--- program second_half_topPaint (robot ABB IRB 5500-27) ---
  Smooth(1)
  Set speed (1000.0 mm/s)
  Set Ref.: FrameTopPaint
  Set Tool: Paint gun
  Show Paint gun
  MoveJ 1 to (-680.86, -907.35, 967.38) mm, rotated rx -105.87 ry 21.86 rz 12.34 deg; joints [-6.464, -4.331, 30.186, -24.09, 51.501, -71.972, -33.04]
  MoveL 2 to (-680.86, -907.35, 967.38) mm, rotated rx -105.87 ry 21.86 rz 12.34 deg; joints [-6.464, -4.331, 30.186, -24.09, 51.501, -71.972, -33.04]
  MoveL 3 to (-711.37, -815.56, 942.01) mm, rotated rx -105.87 ry 21.86 rz 12.34 deg; joints [-10.668, -3.752, 30.735, -25.583, 48.262, -68.348, -33.04]
  MoveL 4 to (-711.37, -815.56, 942.01) mm, rotated rx -105.87 ry 21.86 rz 12.34 deg; joints [-10.668, -3.752, 30.735, -25.583, 48.262, -68.348, -33.04]
  Set speed (50.0 mm/s)
  MoveL 5 to (-723.88, -815.55, 955.73) mm, rotated rx -113.43 ry 35.95 rz 5.6 deg; joints [-9.665, -1.677, 29.706, -47.736, 72.372, -53.861, -33.04]
  MoveL 6 to (-737.5, -815.56, 968.17) mm, rotated rx -117.99 ry 31.14 rz 6.09 deg; joints [-11, -4.053, 28.612, -30.497, 55.555, -56.043, -33.04]
  MoveL 7 to (-752.19, -815.56, 979.36) mm, rotated rx -123.35 ry 26.63 rz 6.68 deg; joints [-13.045, -6.077, 27.151, -7.256, 36.064, -62.575, -33.04]
  MoveL 8 to (-767.89, -815.56, 989.32) mm, rotated rx -137.44 ry 37.1 rz -8.5 deg; joints [-11.723, -3.945, 24.767, -26.574, 60.815, -46.836, -33.04]
  MoveL 9 to (-784.28, -815.56, 997.94) mm, rotated rx -143.37 ry 31.77 rz -8.88 deg; joints [-14.072, -5.42, 22.852, -4.109, 43.017, -52.262, -33.04]
  MoveL 10 to (-800.88, -815.56, 1005.13) mm, rotated rx -160.16 ry 35.48 rz -30.34 deg; joints [-12.936, -2.465, 18.781, -17.366, 67.621, -42.158, -33.04]
  MoveL 11 to (-817.93, -815.56, 1011.14) mm, rotated rx -163.51 ry 29.4 rz -30.19 deg; joints [-15.139, -2.909, 16.546, 0.625, 55.012, -47.084, -33.04]
  MoveL 12 to (-835.41, -815.56, 1016.08) mm, rotated rx -166.27 ry 23.89 rz -30.04 deg; joints [-17.301, -2.699, 14.273, 18.529, 44.337, -54.274, -33.04]
  MoveL 13 to (-853.23, -815.56, 1019.98) mm, rotated rx -168.26 ry 19.06 rz -29.89 deg; joints [-19.167, -1.967, 12.063, 35.166, 36.001, -62.757, -33.04]
  MoveL 14 to (-876.49, -815.56, 1023.58) mm, rotated rx -175.04 ry 16.66 rz -50.25 deg; joints [-17.559, 3.114, 5.489, 8.811, 70.793, -51.29, -33.04]
  MoveL 15 to (-899.83, -815.56, 1025.72) mm, rotated rx -173.61 ry 13.04 rz -49.71 deg; joints [-18.535, 4.811, 2.72, 14.774, 69.055, -56.135, -33.04]
  MoveL 16 to (-923.23, -815.56, 1026.54) mm, rotated rx -171.44 ry 10.87 rz -49.25 deg; joints [-18.954, 6.702, 0.191, 17.247, 69.288, -60.212, -33.04]
  MoveL 17 to (-946.69, -815.56, 1026.19) mm, rotated rx -168.63 ry 9.9 rz -48.73 deg; joints [-18.93, 8.673, -2.078, 17.142, 70.618, -63.617, -33.04]
  MoveL 18 to (-970.21, -815.56, 1024.77) mm, rotated rx -165.25 ry 9.92 rz -48.01 deg; joints [-18.58, 10.662, -4.07, 15.251, 72.434, -66.538, -33.04]
  MoveL 19 to (-993.66, -815.56, 1022.37) mm, rotated rx -161.4 ry 10.72 rz -47 deg; joints [-18.006, 12.618, -5.747, 12.177, 74.323, -69.099, -33.04]
  MoveL 20 to (-1016.91, -815.56, 1019.13) mm, rotated rx -154.6 ry 3.88 rz -27.21 deg; joints [-20.046, 11.059, -3.932, 50.238, 41.644, -92.598, -33.04]
  MoveL 21 to (-1052.97, -815.56, 1012.53) mm, rotated rx -147.18 ry 4.39 rz -25.42 deg; joints [-18.692, 13.832, -5.844, 42.524, 45.231, -94.781, -33.04]
  MoveL 22 to (-1088.6, -815.56, 1004.28) mm, rotated rx -139.61 ry 5.07 rz -23.14 deg; joints [-17.477, 16.361, -7.122, 35.707, 47.402, -97.128, -33.04]
  MoveL 23 to (-1123.86, -815.56, 994.58) mm, rotated rx -132.39 ry 5.54 rz -20.58 deg; joints [-16.529, 18.641, -7.948, 30.174, 48.333, -99.549, -33.04]
  MoveL 24 to (-1158.78, -815.56, 983.54) mm, rotated rx -125.85 ry 5.63 rz -17.99 deg; joints [-15.878, 20.702, -8.533, 26.043, 48.294, -101.998, -33.04]
  MoveL 25 to (-1193.38, -815.56, 971.26) mm, rotated rx -120.15 ry 5.32 rz -15.55 deg; joints [-15.49, 22.587, -9.043, 23.251, 47.542, -104.469, -33.04]
  MoveL 26 to (-1227.05, -815.55, 958.05) mm, rotated rx -117.54 ry 22.59 rz -22.51 deg; joints [-13.683, 27.315, -10.358, -19.064, 74.787, -84.054, -33.04]
  MoveL 27 to (-1260.34, -815.56, 943.78) mm, rotated rx -113.27 ry 22.78 rz -19.28 deg; joints [-13.733, 28.84, -10.662, -21.178, 73.313, -84.803, -33.04]
  MoveL 28 to (-1293.64, -815.56, 929.57) mm, rotated rx -110.3 ry 24.42 rz -16.76 deg; joints [-13.802, 30.363, -10.975, -25.489, 73.688, -83.558, -33.04]
  MoveL 29 to (-1326.93, -815.55, 915.36) mm, rotated rx -110.75 ry 26.95 rz -16.83 deg; joints [-13.938, 32.012, -12.325, -29.467, 76.004, -81.006, -33.04]
  Set speed (1000.0 mm/s)
  MoveL 30 to (-1326.93, -815.55, 915.36) mm, rotated rx -110.75 ry 26.95 rz -16.83 deg; joints [-13.938, 32.012, -12.325, -29.467, 76.004, -81.006, -33.04]
  MoveL 31 to (-1338.64, -909.72, 946.94) mm, rotated rx -108.61 ry 8.09 rz -9.79 deg; joints [-12.86, 29.886, -14.209, 10.126, 49.766, -104.847, -33.04]
  Set speed (1000.0 mm/s)
  MoveL 32 to (-1427.54, -801.91, 1165.8) mm, rotated rx -168.37 ry 26.91 rz -49.4 deg; joints [-18.397, 27.533, -26.297, -2.238, 74.394, -59.791, -33.04]
  MoveL 33 to (-1441.08, -755.13, 1078.46) mm, rotated rx -168.37 ry 26.91 rz -49.4 deg; joints [-19.651, 28.149, -23.955, -2.229, 72.544, -56.455, -33.04]
  MoveL 34 to (-1441.08, -755.13, 1078.46) mm, rotated rx -168.37 ry 26.91 rz -49.4 deg; joints [-19.651, 28.149, -23.955, -2.229, 72.544, -56.455, -33.04]
  Set speed (50.0 mm/s)
  MoveL 35 to (-1392.85, -755.13, 1070.73) mm, rotated rx -167.45 ry 26.52 rz -49.02 deg; joints [-19.416, 26.202, -21.042, -2.719, 73.023, -56.398, -33.04]
  MoveL 36 to (-1344.51, -755.13, 1064.62) mm, rotated rx -166.39 ry 26.02 rz -48.59 deg; joints [-19.179, 24.323, -18.348, -2.991, 73.454, -56.694, -33.04]
  MoveL 37 to (-1296.05, -755.13, 1060.31) mm, rotated rx -165.14 ry 25.36 rz -48.07 deg; joints [-18.944, 22.516, -15.888, -2.97, 73.811, -57.435, -33.04]
  MoveL 38 to (-1247.5, -755.13, 1057.45) mm, rotated rx -163.92 ry 24.63 rz -47.58 deg; joints [-18.714, 20.718, -13.548, -2.801, 74.124, -58.304, -33.04]
  MoveL 39 to (-1198.88, -755.13, 1055.53) mm, rotated rx -162.66 ry 23.79 rz -47.07 deg; joints [-18.49, 18.954, -11.35, -2.42, 74.383, -59.409, -33.04]
  MoveL 40 to (-1154.65, -755.13, 1054.25) mm, rotated rx -161.47 ry 22.9 rz -46.6 deg; joints [-18.296, 17.383, -9.469, -1.877, 74.573, -60.622, -33.04]
  MoveL 41 to (-1110.41, -755.13, 1053.12) mm, rotated rx -160.23 ry 21.86 rz -46.13 deg; joints [-18.116, 15.849, -7.702, -1.119, 74.72, -62.054, -33.04]
  MoveL 42 to (-1066.18, -755.13, 1051.84) mm, rotated rx -158.93 ry 20.61 rz -45.66 deg; joints [-17.96, 14.367, -6.063, -0.094, 74.823, -63.754, -33.04]
  MoveL 43 to (-1021.98, -755.13, 1050.14) mm, rotated rx -155.56 ry 16.38 rz -27.11 deg; joints [-20.211, 7.807, 1.212, 35.102, 38.519, -76.601, -33.04]
  MoveL 44 to (-977.83, -755.13, 1047.71) mm, rotated rx -167.34 ry 20.31 rz -48.51 deg; joints [-18.414, 8.637, -0.031, 2.711, 72.736, -56.241, -33.04]
  MoveL 45 to (-933.79, -755.13, 1044.23) mm, rotated rx -172.03 ry 17.59 rz -49.64 deg; joints [-19.417, 5.728, 2.312, 9.306, 68.998, -54.431, -33.04]
  MoveL 46 to (-889.96, -755.13, 1039.39) mm, rotated rx -176.35 ry 15.79 rz -50.43 deg; joints [-20.284, 2.79, 5.029, 14.554, 65.44, -52.144, -33.04]
  MoveL 47 to (-859.98, -755.13, 1035.09) mm, rotated rx -179.05 ry 15.23 rz -50.85 deg; joints [-20.714, 0.773, 7.104, 16.981, 63.333, -50.184, -33.04]
  MoveL 48 to (-830.15, -755.13, 1029.86) mm, rotated rx 178.5 ry 15.31 rz -51.25 deg; joints [-20.935, -1.226, 9.339, 18.054, 61.765, -47.765, -33.04]
  MoveL 49 to (-800.49, -755.13, 1023.59) mm, rotated rx 176.32 ry 16.12 rz -51.7 deg; joints [-20.879, -3.182, 11.724, 17.357, 61.061, -44.748, -33.04]
  MoveL 50 to (-771.02, -755.13, 1016.11) mm, rotated rx 174.42 ry 17.73 rz -52.29 deg; joints [-20.476, -5.053, 14.244, 14.483, 61.629, -41.047, -33.04]
  MoveL 51 to (-746.27, -755.13, 1008.74) mm, rotated rx 173.04 ry 19.75 rz -52.97 deg; joints [-19.815, -6.52, 16.467, 10.081, 63.46, -37.399, -33.04]
  MoveL 52 to (-721.93, -755.13, 1000.39) mm, rotated rx 171.85 ry 22.37 rz -53.89 deg; joints [-18.839, -7.804, 18.74, 3.824, 66.801, -33.461, -33.04]
  MoveL 53 to (-698.07, -755.13, 991) mm, rotated rx 170.81 ry 25.58 rz -55.13 deg; joints [-17.554, -8.832, 21.041, -4.204, 71.863, -29.519, -33.04]
  MoveL 54 to (-674.71, -755.13, 980.5) mm, rotated rx -178.47 ry 30.85 rz -33.67 deg; joints [-19.518, -13.327, 26.774, 8.833, 42.793, -34.507, -33.04]
  MoveL 55 to (-651.88, -755.13, 968.81) mm, rotated rx -177.42 ry 35.05 rz -34.68 deg; joints [-17.437, -13.741, 29.013, -6.651, 53.844, -28.419, -33.04]
  MoveL 56 to (-629.61, -755.13, 955.87) mm, rotated rx -176.18 ry 39.58 rz -35.92 deg; joints [-15.275, -13.645, 31.207, -21.324, 65.847, -24.476, -33.04]
  MoveL 57 to (-609.19, -755.13, 942.47) mm, rotated rx -157.46 ry 39.23 rz -11.27 deg; joints [-17.521, -17.024, 35.308, -13.254, 41.312, -30.381, -33.04]
  MoveL 58 to (-589.56, -755.13, 927.98) mm, rotated rx -153.88 ry 43.02 rz -11.42 deg; joints [-15.133, -16.253, 37.231, -29.816, 56.214, -26.857, -33.04]
  MoveL 59 to (-570.79, -755.13, 912.43) mm, rotated rx -150.35 ry 46.8 rz -11.58 deg; joints [-13.086, -14.971, 38.921, -43.447, 70.123, -26.03, -33.04]
  MoveL 60 to (-552.87, -755.13, 895.83) mm, rotated rx -132.12 ry 37.38 rz 9.39 deg; joints [-15.418, -17.926, 41.46, -31.974, 44.911, -34.545, -33.04]
  MoveL 61 to (-535.98, -755.13, 878.3) mm, rotated rx -128.2 ry 40.11 rz 9.17 deg; joints [-13.411, -16.317, 42.937, -45.251, 59.152, -33.515, -33.04]
  MoveL 62 to (-519.26, -755.12, 858.88) mm, rotated rx -124.45 ry 42.99 rz 8.96 deg; joints [-11.739, -14.257, 44.196, -56.795, 72.787, -34.124, -33.04]
  MoveL 63 to (-503.73, -755.13, 838.65) mm, rotated rx -114.08 ry 28.02 rz 20.35 deg; joints [-13.853, -17.337, 45.471, -36.435, 43.409, -46.335, -33.04]
  MoveL 64 to (-489.34, -755.13, 817.63) mm, rotated rx -111.22 ry 30.33 rz 19.47 deg; joints [-12.23, -15.335, 46.617, -48.302, 56.678, -44.847, -33.04]
  MoveL 65 to (-476.03, -755.13, 795.85) mm, rotated rx -108.72 ry 32.65 rz 18.71 deg; joints [-10.971, -13.136, 47.527, -57.964, 68.476, -44.674, -33.04]
  MoveL 66 to (-463.75, -755.13, 773.36) mm, rotated rx -104.02 ry 15.61 rz 23.88 deg; joints [-13.073, -16.444, 47.716, -24.573, 33.094, -63.727, -33.04]
  MoveL 67 to (-452.46, -755.13, 750.19) mm, rotated rx -102.19 ry 17.65 rz 22.76 deg; joints [-11.641, -14.473, 48.652, -37.695, 45.898, -59.342, -33.04]
  Set speed (1000.0 mm/s)
  MoveL 68 to (-452.46, -755.13, 750.19) mm, rotated rx -102.19 ry 17.65 rz 22.76 deg; joints [-11.641, -14.473, 48.652, -37.695, 45.898, -59.342, -33.04]
  MoveL 69 to (-408.75, -842.79, 770.31) mm, rotated rx -102.19 ry 17.65 rz 22.76 deg; joints [-5.982, -16.094, 48.843, -32.575, 47.942, -65.004, -33.04]
  Set speed (1000.0 mm/s)
  MoveL 70 to (-280.85, -767.56, 751.15) mm, rotated rx -114.97 ry 33.92 rz 24.38 deg; joints [-10.377, -28.704, 57.94, -50.266, 54.482, -37.789, -33.04]
  MoveL 71 to (-339.72, -694.7, 716.13) mm, rotated rx -114.97 ry 33.92 rz 24.38 deg; joints [-16.491, -24.096, 57.105, -61.18, 58.103, -29.538, -33.04]
  MoveL 72 to (-339.72, -694.7, 716.13) mm, rotated rx -114.97 ry 33.92 rz 24.38 deg; joints [-16.491, -24.096, 57.105, -61.18, 58.103, -29.538, -33.04]
  Set speed (50.0 mm/s)
  MoveL 73 to (-357.11, -694.7, 743.86) mm, rotated rx -117.94 ry 32.09 rz 25.15 deg; joints [-18.606, -26.389, 55.654, -51.693, 45.003, -28.551, -33.04]
  MoveL 74 to (-375.74, -694.69, 770.58) mm, rotated rx -130.67 ry 46.61 rz 11.02 deg; joints [-15.598, -23.039, 54.114, -63.974, 72.081, -20.66, -33.04]
  MoveL 75 to (-395.64, -694.7, 796.31) mm, rotated rx -134.35 ry 44.15 rz 11.08 deg; joints [-17.761, -25.145, 52.527, -53.816, 58.424, -18.794, -33.04]
  MoveL 76 to (-416.85, -694.7, 820.98) mm, rotated rx -138.3 ry 41.66 rz 11.13 deg; joints [-20.283, -26.646, 50.605, -42.162, 44.019, -18.14, -33.04]
  MoveL 77 to (-439.4, -694.7, 844.57) mm, rotated rx -159.64 ry 49.05 rz -13.25 deg; joints [-17.084, -23.648, 47.731, -45.094, 65.338, -13.723, -33.04]
  MoveL 78 to (-462.87, -694.7, 866.64) mm, rotated rx -162.58 ry 45.48 rz -12.83 deg; joints [-19.593, -24.599, 45.602, -31.764, 50.861, -14.485, -33.04]
  MoveL 79 to (-487.43, -694.7, 887.42) mm, rotated rx 175.77 ry 43.79 rz -39.75 deg; joints [-16.92, -21.228, 41.257, -31.131, 70.359, -12.811, -33.04]
  MoveL 80 to (-513.03, -694.7, 906.91) mm, rotated rx 175.37 ry 39.79 rz -37.93 deg; joints [-19.194, -21.396, 38.943, -17.947, 57.935, -15.44, -33.04]
  MoveL 81 to (-539.61, -694.7, 925.1) mm, rotated rx 174.96 ry 35.98 rz -36.42 deg; joints [-21.423, -21.016, 36.518, -3.67, 46.106, -20.168, -33.04]
  MoveL 82 to (-567.52, -694.7, 942.26) mm, rotated rx 162.99 ry 28.48 rz -57.97 deg; joints [-19.195, -16.589, 30.728, -8.728, 70.789, -18.654, -33.04]
  MoveL 83 to (-596.05, -694.71, 958.02) mm, rotated rx 164.29 ry 25.51 rz -56.36 deg; joints [-20.66, -15.521, 28.236, -0.029, 64.448, -22.61, -33.04]
  MoveL 84 to (-625.13, -694.71, 972.48) mm, rotated rx 165.62 ry 23.02 rz -55.12 deg; joints [-21.799, -14.167, 25.764, 7.202, 59.845, -26.748, -33.04]
  MoveL 85 to (-654.73, -694.71, 985.73) mm, rotated rx 167.01 ry 21.02 rz -54.2 deg; joints [-22.603, -12.611, 23.335, 12.74, 56.867, -30.707, -33.04]
  MoveL 86 to (-684.8, -694.71, 997.88) mm, rotated rx 168.52 ry 19.53 rz -53.53 deg; joints [-23.088, -10.915, 20.962, 16.48, 55.343, -34.23, -33.04]
  MoveL 87 to (-715.3, -694.71, 1009.03) mm, rotated rx 170.16 ry 18.56 rz -53.05 deg; joints [-23.288, -9.129, 18.656, 18.478, 55.039, -37.199, -33.04]
  MoveL 88 to (-746.19, -694.71, 1019.28) mm, rotated rx 171.94 ry 18.1 rz -52.71 deg; joints [-23.247, -7.286, 16.425, 18.902, 55.71, -39.601, -33.04]
  MoveL 89 to (-790.01, -694.71, 1032.3) mm, rotated rx 171.82 ry 18.31 rz -52.78 deg; joints [-23.382, -5.469, 14.353, 18.926, 55.572, -39.688, -33.04]
  MoveL 90 to (-834.27, -694.71, 1044) mm, rotated rx -164.38 ry 12.66 rz -47.66 deg; joints [-21.172, 3.673, 3.763, 15.498, 67.78, -65.474, -33.04]
  MoveL 91 to (-878.76, -694.71, 1054.62) mm, rotated rx -165.86 ry 14.3 rz -47.99 deg; joints [-21.21, 4.9, 2.353, 14.26, 67.353, -63.309, -33.04]
  MoveL 92 to (-923.43, -694.71, 1064.45) mm, rotated rx -167.05 ry 15.38 rz -48.3 deg; joints [-21.336, 6.309, 0.654, 13.66, 66.935, -61.91, -33.04]
  MoveL 93 to (-968.22, -694.71, 1073.75) mm, rotated rx -168.04 ry 16.15 rz -48.56 deg; joints [-21.499, 7.83, -1.235, 13.422, 66.525, -60.996, -33.04]
  MoveL 94 to (-1026.95, -694.71, 1085.57) mm, rotated rx -169.1 ry 16.87 rz -48.86 deg; joints [-21.736, 9.93, -3.917, 13.442, 66.008, -60.295, -33.04]
  MoveL 95 to (-1085.65, -694.71, 1097.49) mm, rotated rx -170.03 ry 17.43 rz -49.12 deg; joints [-21.979, 12.104, -6.785, 13.695, 65.517, -59.971, -33.04]
  MoveL 96 to (-1144.22, -694.71, 1110.04) mm, rotated rx -170.86 ry 17.87 rz -49.36 deg; joints [-22.222, 14.329, -9.82, 14.113, 65.054, -59.935, -33.04]
  MoveL 97 to (-1179.59, -694.71, 1109.54) mm, rotated rx -170.86 ry 17.87 rz -49.36 deg; joints [-22.351, 15.89, -11.706, 14.449, 64.884, -60.342, -33.04]
  MoveL 98 to (-1214.81, -694.71, 1107.82) mm, rotated rx -170.86 ry 17.87 rz -49.36 deg; joints [-22.474, 17.461, -13.593, 14.773, 64.725, -60.738, -33.04]
  MoveL 99 to (-1249.9, -694.71, 1104.91) mm, rotated rx -170.86 ry 17.87 rz -49.36 deg; joints [-22.592, 19.043, -15.485, 15.086, 64.575, -61.127, -33.04]
  MoveL 100 to (-1284.86, -694.71, 1100.85) mm, rotated rx -170.86 ry 17.87 rz -49.36 deg; joints [-22.705, 20.637, -17.385, 15.39, 64.435, -61.509, -33.04]
  MoveL 101 to (-1321.33, -694.71, 1095.39) mm, rotated rx -170.86 ry 17.87 rz -49.36 deg; joints [-22.819, 22.322, -19.388, 15.7, 64.298, -61.906, -33.04]
  MoveL 102 to (-1357.66, -694.71, 1088.73) mm, rotated rx -170.86 ry 17.87 rz -49.36 deg; joints [-22.928, 24.024, -21.407, 16.001, 64.172, -62.301, -33.04]
  MoveL 103 to (-1393.86, -694.71, 1080.88) mm, rotated rx -170.86 ry 17.87 rz -49.36 deg; joints [-23.032, 25.746, -23.447, 16.297, 64.055, -62.698, -33.04]
  Set speed (1000.0 mm/s)
  MoveL 104 to (-1393.86, -694.71, 1080.88) mm, rotated rx -170.86 ry 17.87 rz -49.36 deg; joints [-23.032, 25.746, -23.447, 16.297, 64.055, -62.698, -33.04]
  MoveL 105 to (-1386.19, -728.04, 1174.85) mm, rotated rx -170.86 ry 17.87 rz -49.36 deg; joints [-22.138, 25.351, -26.342, 16.111, 66.402, -66.107, -33.04]
  Set speed (1000.0 mm/s)
  MoveL 106 to (-1383.57, -648.28, 1177.84) mm, rotated rx -164.63 ry -10.56 rz -30.24 deg; joints [-29.593, 31.056, -38.749, 68.964, 56.594, -115.064, -33.04]
  MoveL 107 to (-1354.96, -634.29, 1083.04) mm, rotated rx -162.02 ry -4.77 rz -49.56 deg; joints [-27.513, 32.255, -36.738, 33.77, 75.893, -92.359, -33.04]
  MoveL 108 to (-1354.96, -634.29, 1083.04) mm, rotated rx -162.02 ry -4.77 rz -49.56 deg; joints [-27.513, 32.255, -36.738, 33.77, 75.893, -92.359, -33.04]
  Set speed (50.0 mm/s)
  MoveL 109 to (-1316.03, -634.28, 1090.58) mm, rotated rx -162.02 ry -4.77 rz -49.56 deg; joints [-27.496, 30.204, -34.071, 34.005, 75.314, -91.786, -33.04]
  MoveL 110 to (-1276.87, -634.28, 1096.8) mm, rotated rx -164.09 ry -4.88 rz -49.8 deg; joints [-27.831, 27.6, -30.819, 36.058, 73.417, -89.721, -33.04]
  MoveL 111 to (-1237.63, -634.28, 1101.65) mm, rotated rx -166.2 ry -4.97 rz -49.99 deg; joints [-28.188, 25.02, -27.61, 38.256, 71.356, -87.707, -33.04]
  MoveL 112 to (-1198.44, -634.28, 1105.09) mm, rotated rx -168.35 ry -5.02 rz -50.12 deg; joints [-28.564, 22.461, -24.431, 40.594, 69.113, -85.742, -33.04]
  MoveL 113 to (-1159.29, -634.28, 1107.12) mm, rotated rx -170.59 ry -4.99 rz -50.21 deg; joints [-28.959, 19.891, -21.234, 43.1, 66.607, -83.778, -33.04]
  MoveL 114 to (-1117.81, -634.28, 1107.7) mm, rotated rx -172.95 ry -4.89 rz -50.24 deg; joints [-29.388, 17.188, -17.865, 45.87, 63.758, -81.788, -33.04]
  MoveL 115 to (-1076.38, -634.28, 1106.64) mm, rotated rx -175.36 ry -4.66 rz -50.22 deg; joints [-29.827, 14.475, -14.468, 48.789, 60.627, -79.838, -33.04]
  MoveL 116 to (-1035, -634.28, 1103.91) mm, rotated rx -177.81 ry -4.29 rz -50.16 deg; joints [-30.273, 11.746, -11.032, 51.858, 57.195, -77.929, -33.04]
  MoveL 117 to (-993.67, -634.28, 1099.48) mm, rotated rx 179.68 ry -3.75 rz -50.05 deg; joints [-30.726, 8.988, -7.535, 55.102, 53.417, -76.051, -33.04]
  MoveL 118 to (-952.39, -634.28, 1093.3) mm, rotated rx 177.08 ry -3.02 rz -49.91 deg; joints [-31.187, 6.183, -3.95, 58.575, 49.223, -74.195, -33.04]
  MoveL 119 to (-911.16, -634.28, 1085.32) mm, rotated rx 170.97 ry -0.42 rz -49.61 deg; joints [-32.081, 1.909, 1.768, 66.623, 38.914, -70.262, -33.04]
  MoveL 120 to (-870.06, -634.28, 1072.26) mm, rotated rx 161.64 ry 24.15 rz -56.14 deg; joints [-25.915, -5.114, 14.971, 12.913, 51.726, -25.277, -33.04]
  MoveL 121 to (-829.03, -634.28, 1058.97) mm, rotated rx 161.64 ry 24.15 rz -56.14 deg; joints [-25.807, -6.839, 17.044, 12.396, 52.013, -24.786, -33.04]
  MoveL 122 to (-788.13, -634.28, 1045.27) mm, rotated rx 161.64 ry 24.15 rz -56.14 deg; joints [-25.693, -8.569, 19.094, 11.9, 52.305, -24.332, -33.04]
  MoveL 123 to (-747.44, -634.28, 1031) mm, rotated rx 161.64 ry 24.15 rz -56.14 deg; joints [-25.573, -10.301, 21.124, 11.421, 52.602, -23.909, -33.04]
  MoveL 124 to (-707.08, -634.28, 1015.99) mm, rotated rx 161.64 ry 24.15 rz -56.14 deg; joints [-25.446, -12.03, 23.135, 10.949, 52.909, -23.506, -33.04]
  MoveL 125 to (-667.17, -634.28, 1000.09) mm, rotated rx 161.64 ry 24.15 rz -56.14 deg; joints [-25.312, -13.749, 25.129, 10.477, 53.228, -23.113, -33.04]
  MoveL 126 to (-627.79, -634.28, 983.13) mm, rotated rx 161.64 ry 24.15 rz -56.14 deg; joints [-25.169, -15.454, 27.11, 9.996, 53.562, -22.721, -33.04]
  MoveL 127 to (-589.03, -634.28, 964.94) mm, rotated rx 161.64 ry 24.15 rz -56.14 deg; joints [-25.018, -17.14, 29.081, 9.495, 53.916, -22.317, -33.04]
  MoveL 128 to (-521.38, -634.28, 928.72) mm, rotated rx 160.54 ry 25.2 rz -56.78 deg; joints [-24.397, -20.285, 33.162, 5.492, 56.262, -19.182, -33.04]
  MoveL 129 to (-488.54, -634.28, 908.62) mm, rotated rx 159.09 ry 27.55 rz -58.21 deg; joints [-23.17, -21.751, 35.826, -2.329, 61.681, -14.851, -33.04]
  MoveL 130 to (-456.44, -634.28, 887.04) mm, rotated rx 157.59 ry 30.29 rz -60.07 deg; joints [-21.582, -22.904, 38.513, -11.425, 68.849, -10.813, -33.04]
  MoveL 131 to (-425.22, -634.28, 863.92) mm, rotated rx 170.2 ry 39.25 rz -38.62 deg; joints [-24.275, -27.281, 44.353, -11.924, 47.46, -10, -33.04]
  MoveL 132 to (-397.94, -634.28, 841.74) mm, rotated rx 170.15 ry 42.47 rz -40.29 deg; joints [-22.129, -27.683, 46.769, -24.269, 58.676, -6.356, -33.04]
  MoveL 133 to (-371.77, -634.27, 818.47) mm, rotated rx 170.03 ry 45.79 rz -42.27 deg; joints [-19.915, -27.569, 49.069, -35.693, 70.343, -4.4, -33.04]
  MoveL 134 to (-346.75, -634.28, 794.12) mm, rotated rx -166.97 ry 48.65 rz -13.97 deg; joints [-23.649, -30.931, 53.337, -40.952, 52.991, -3.509, -33.04]
  MoveL 135 to (-322.86, -634.28, 768.67) mm, rotated rx -164.78 ry 51.68 rz -14.53 deg; joints [-21.227, -30.129, 55.493, -51.709, 65.924, -3.715, -33.04]
  MoveL 136 to (-300.1, -634.28, 742.13) mm, rotated rx -141.36 ry 45.05 rz 12.36 deg; joints [-25.779, -33.162, 58.341, -56.228, 47.993, -3.726, -33.04]
  MoveL 137 to (-278.48, -634.28, 714.5) mm, rotated rx -137.94 ry 47.13 rz 12.43 deg; joints [-23.334, -31.875, 60.333, -64.364, 60.071, -6.057, -33.04]
  MoveL 138 to (-257.97, -634.28, 685.8) mm, rotated rx -123.43 ry 33.52 rz 29.26 deg; joints [-27.848, -34.937, 61.807, -64.029, 38.79, -8.276, -33.04]
  Set speed (1000.0 mm/s)
  MoveL 139 to (-257.97, -634.28, 685.8) mm, rotated rx -123.43 ry 33.52 rz 29.26 deg; joints [-27.848, -34.937, 61.807, -64.029, 38.79, -8.276, -33.04]
  MoveL 140 to (-190.63, -692.21, 731.73) mm, rotated rx -134.65 ry 49.19 rz 12.51 deg; joints [-15.298, -37.261, 63.293, -59.641, 65.012, -17.041, -33.04]
  Set speed (1000.0 mm/s)
  MoveL 141 to (-122.9, -618.87, 712.66) mm, rotated rx -142.88 ry 47.91 rz 13.38 deg; joints [-29.119, -48.176, 66.475, -50.842, 38.175, -0.586, -33.04]
  MoveL 142 to (-194.43, -573.85, 659.22) mm, rotated rx -142.88 ry 47.91 rz 13.38 deg; joints [-32.599, -38.02, 65.244, -72.969, 55.346, 9.693, -33.04]
  MoveL 143 to (-194.43, -573.85, 659.22) mm, rotated rx -142.88 ry 47.91 rz 13.38 deg; joints [-32.599, -38.02, 65.244, -72.969, 55.346, 9.693, -33.04]
  Set speed (50.0 mm/s)
  MoveL 144 to (-219.42, -573.85, 691.19) mm, rotated rx -168.5 ry 53.82 rz -15.6 deg; joints [-26.592, -35.485, 62.253, -59.133, 66.795, 5.859, -33.04]
  MoveL 145 to (-245.66, -573.85, 721.92) mm, rotated rx -170.35 ry 50.93 rz -14.9 deg; joints [-29.075, -36.259, 59.872, -49.532, 54.056, 6.877, -33.04]
  MoveL 146 to (-273.13, -573.85, 751.4) mm, rotated rx 165.69 ry 46.89 rz -44 deg; joints [-24.248, -33.143, 55.523, -38.026, 67.49, 3.047, -33.04]
  MoveL 147 to (-301.84, -573.85, 779.65) mm, rotated rx 166.16 ry 43.83 rz -41.85 deg; joints [-26.546, -33.105, 53.003, -26.934, 55.657, 1.11, -33.04]
  MoveL 148 to (-331.74, -573.84, 806.69) mm, rotated rx 152.1 ry 33.68 rz -63.59 deg; joints [-23.32, -29.086, 47.36, -20.418, 72.694, -1.696, -33.04]
  MoveL 149 to (-362.3, -573.85, 832.06) mm, rotated rx 153.68 ry 31.23 rz -61.45 deg; joints [-25.042, -28.271, 44.813, -11.519, 64.603, -4.897, -33.04]
  MoveL 150 to (-393.95, -573.85, 856.32) mm, rotated rx 155.14 ry 28.97 rz -59.69 deg; joints [-26.496, -27.094, 42.224, -3.137, 57.77, -8.726, -33.04]
  MoveL 151 to (-426.44, -573.85, 879.33) mm, rotated rx 155.14 ry 28.97 rz -59.69 deg; joints [-26.613, -25.628, 40.437, -2.635, 57.395, -9.123, -33.04]
  MoveL 152 to (-459.61, -573.85, 901.11) mm, rotated rx 155.14 ry 28.97 rz -59.69 deg; joints [-26.721, -24.133, 38.65, -2.172, 57.051, -9.487, -33.04]
  MoveL 153 to (-499.91, -573.85, 925.56) mm, rotated rx 155.14 ry 28.97 rz -59.69 deg; joints [-26.84, -22.326, 36.52, -1.659, 56.673, -9.893, -33.04]
  MoveL 154 to (-541.01, -573.85, 948.56) mm, rotated rx 155.14 ry 28.97 rz -59.69 deg; joints [-26.95, -20.496, 34.383, -1.173, 56.32, -10.28, -33.04]
  MoveL 155 to (-582.81, -573.85, 970.29) mm, rotated rx 155.14 ry 28.97 rz -59.69 deg; joints [-27.051, -18.65, 32.237, -0.7, 55.985, -10.662, -33.04]
  MoveL 156 to (-625.21, -573.85, 990.93) mm, rotated rx 155.14 ry 28.97 rz -59.69 deg; joints [-27.145, -16.796, 30.078, -0.227, 55.66, -11.054, -33.04]
  MoveL 157 to (-668.11, -573.85, 1010.65) mm, rotated rx 155.14 ry 28.97 rz -59.69 deg; joints [-27.234, -14.939, 27.903, 0.257, 55.338, -11.465, -33.04]
  MoveL 158 to (-711.41, -573.85, 1029.64) mm, rotated rx 155.14 ry 28.97 rz -59.69 deg; joints [-27.317, -13.084, 25.708, 0.764, 55.014, -11.906, -33.04]
  MoveL 159 to (-748.06, -573.85, 1043.66) mm, rotated rx 157.61 ry 6.44 rz -70.97 deg; joints [-30.214, -6.982, 13.644, 24.862, 64.48, -31.395, -33.04]
  MoveL 160 to (-785.01, -573.85, 1056.24) mm, rotated rx 159.54 ry 6.06 rz -70.87 deg; joints [-30.059, -4.756, 10.809, 24.468, 66.213, -33.972, -33.04]
  MoveL 161 to (-822.27, -573.85, 1067.4) mm, rotated rx 161.68 ry 5.81 rz -70.82 deg; joints [-29.825, -2.438, 7.89, 23.534, 68.351, -36.593, -33.04]
  MoveL 162 to (-859.82, -573.85, 1077.12) mm, rotated rx 163.93 ry 5.7 rz -70.8 deg; joints [-29.537, -0.058, 4.925, 22.194, 70.729, -39.212, -33.04]
  MoveL 163 to (-897.67, -573.85, 1085.42) mm, rotated rx 166.26 ry 5.73 rz -70.79 deg; joints [-29.212, 2.369, 1.93, 20.532, 73.248, -41.818, -33.04]
  MoveL 164 to (-935.15, -573.85, 1092.2) mm, rotated rx 171.31 ry 9.42 rz -50.91 deg; joints [-31.484, 1.113, 4.075, 53.364, 36.921, -59.511, -33.04]
  MoveL 165 to (-972.91, -573.85, 1097.61) mm, rotated rx 173.72 ry 8.88 rz -50.75 deg; joints [-31.012, 3.518, 1.087, 50.816, 40.223, -61.321, -33.04]
  MoveL 166 to (-1010.95, -573.85, 1101.66) mm, rotated rx 176.22 ry 8.44 rz -50.58 deg; joints [-30.529, 5.963, -1.923, 48.198, 43.461, -63.201, -33.04]
  MoveL 167 to (-1049.28, -573.85, 1104.34) mm, rotated rx 179.02 ry 8.02 rz -50.35 deg; joints [-30.017, 8.52, -5.057, 45.445, 46.81, -65.379, -33.04]
  MoveL 168 to (-1095.21, -573.85, 1105.76) mm, rotated rx 178.6 ry -0.8 rz -49.98 deg; joints [-32.096, 12.453, -11.192, 57.274, 48.606, -75.574, -33.04]
  MoveL 169 to (-1141.03, -573.85, 1105.26) mm, rotated rx -179.95 ry -2.76 rz -50.03 deg; joints [-32.127, 15.498, -15.21, 56.44, 52.134, -78.187, -33.04]
  MoveL 170 to (-1186.71, -573.85, 1102.88) mm, rotated rx -178.47 ry -4.6 rz -50.15 deg; joints [-32.125, 18.597, -19.315, 55.198, 55.858, -80.655, -33.04]
  MoveL 171 to (-1232.24, -573.85, 1098.69) mm, rotated rx -176.96 ry -6.34 rz -50.33 deg; joints [-32.096, 21.761, -23.526, 53.627, 59.732, -83.045, -33.04]
  MoveL 172 to (-1277.62, -573.85, 1092.71) mm, rotated rx -175.43 ry -7.97 rz -50.56 deg; joints [-32.044, 25.002, -27.87, 51.781, 63.733, -85.408, -33.04]
  MoveL 173 to (-1322.87, -573.85, 1084.99) mm, rotated rx -173.88 ry -9.5 rz -50.83 deg; joints [-31.971, 28.336, -32.379, 49.693, 67.845, -87.788, -33.04]
  Set speed (1000.0 mm/s)
  MoveL 174 to (-1322.87, -573.85, 1084.99) mm, rotated rx -173.88 ry -9.5 rz -50.83 deg; joints [-31.971, 28.336, -32.379, 49.693, 67.845, -87.788, -33.04]
  MoveL 175 to (-1341.5, -567.86, 1183.06) mm, rotated rx -173.88 ry -9.5 rz -50.83 deg; joints [-32.09, 29.766, -38.022, 47.112, 72.847, -91.048, -33.04]
  Set speed (1000.0 mm/s)
  MoveL 176 to (-1313.29, -509.41, 1185.2) mm, rotated rx -174 ry -7.96 rz -50.61 deg; joints [-33.45, 27.776, -35.021, 50.071, 68.116, -90.852, -33.04]
  MoveL 177 to (-1296.48, -513.43, 1086.71) mm, rotated rx -174 ry -7.96 rz -50.61 deg; joints [-33.386, 26.559, -29.695, 52.526, 63.238, -87.794, -33.04]
  MoveL 178 to (-1296.48, -513.43, 1086.71) mm, rotated rx -174 ry -7.96 rz -50.61 deg; joints [-33.386, 26.559, -29.695, 52.526, 63.238, -87.794, -33.04]
  Set speed (50.0 mm/s)
  MoveL 179 to (-1258.34, -513.43, 1092.62) mm, rotated rx -175.35 ry -6.81 rz -50.43 deg; joints [-33.519, 23.847, -26.066, 54.385, 59.91, -85.983, -33.04]
  MoveL 180 to (-1220.17, -513.43, 1097.33) mm, rotated rx -176.67 ry -5.59 rz -50.28 deg; joints [-33.643, 21.197, -22.544, 56.13, 56.627, -84.205, -33.04]
  MoveL 181 to (-1182, -513.43, 1100.83) mm, rotated rx -177.98 ry -4.32 rz -50.15 deg; joints [-33.757, 18.6, -19.111, 57.751, 53.389, -82.439, -33.04]
  MoveL 182 to (-1143.81, -513.43, 1103.09) mm, rotated rx -179.27 ry -2.98 rz -50.06 deg; joints [-33.861, 16.049, -15.756, 59.23, 50.207, -80.666, -33.04]
  MoveL 183 to (-1104.9, -513.43, 1104.12) mm, rotated rx 179.43 ry -1.55 rz -50 deg; joints [-33.953, 13.492, -12.406, 60.563, 47.035, -78.826, -33.04]
  MoveL 184 to (-1065.98, -513.43, 1103.84) mm, rotated rx 178.15 ry -0.05 rz -49.98 deg; joints [-34.03, 10.973, -9.113, 61.684, 43.954, -76.92, -33.04]
  MoveL 185 to (-1027.05, -513.43, 1102.23) mm, rotated rx 176.88 ry 1.52 rz -50.02 deg; joints [-34.089, 8.485, -5.869, 62.538, 40.995, -74.907, -33.04]
  MoveL 186 to (-988.09, -513.43, 1099.26) mm, rotated rx 175.63 ry 3.14 rz -50.1 deg; joints [-34.128, 6.029, -2.671, 63.054, 38.21, -72.742, -33.04]
  MoveL 187 to (-949.11, -513.43, 1094.89) mm, rotated rx 173.09 ry 2.63 rz -70.17 deg; joints [-31.467, 7.286, -4.699, 23.829, 75.046, -52.259, -33.04]
  MoveL 188 to (-910.16, -513.43, 1089.13) mm, rotated rx 171.34 ry 3.87 rz -70.35 deg; joints [-31.36, 4.857, -1.509, 23.346, 73.511, -49.275, -33.04]
  MoveL 189 to (-871.59, -513.43, 1081.99) mm, rotated rx 169.6 ry 5.16 rz -70.6 deg; joints [-31.216, 2.485, 1.618, 22.513, 72.252, -46.22, -33.04]
  MoveL 190 to (-833.49, -513.43, 1073.52) mm, rotated rx 170.67 ry 6.91 rz -70.89 deg; joints [-30.503, 1.119, 3.619, 18.651, 74.196, -45.432, -33.04]
  MoveL 191 to (-795.86, -513.42, 1063.72) mm, rotated rx 170.67 ry 6.91 rz -70.89 deg; joints [-30.541, -0.485, 5.598, 18.7, 73.934, -45.052, -33.04]
  MoveL 192 to (-758.7, -513.42, 1052.61) mm, rotated rx 170.67 ry 6.91 rz -70.89 deg; joints [-30.58, -2.064, 7.563, 18.747, 73.667, -44.66, -33.04]
  MoveL 193 to (-719.79, -513.42, 1039.41) mm, rotated rx 170.67 ry 6.91 rz -70.89 deg; joints [-30.622, -3.712, 9.635, 18.794, 73.376, -44.23, -33.04]
  MoveL 194 to (-681.4, -513.42, 1024.77) mm, rotated rx 149.35 ry 33.54 rz -64.1 deg; joints [-28.786, -14.613, 29.431, -12.165, 61.244, -1.134, -33.04]
  MoveL 195 to (-643.51, -513.42, 1008.71) mm, rotated rx 149.35 ry 33.54 rz -64.1 deg; joints [-28.764, -16.254, 31.317, -12.486, 61.457, -0.85, -33.04]
  MoveL 196 to (-606.12, -513.42, 991.24) mm, rotated rx 149.35 ry 33.54 rz -64.1 deg; joints [-28.739, -17.877, 33.204, -12.834, 61.689, -0.544, -33.04]
  MoveL 197 to (-569.22, -513.42, 972.38) mm, rotated rx 149.35 ry 33.54 rz -64.1 deg; joints [-28.71, -19.483, 35.094, -13.21, 61.943, -0.217, -33.04]
  MoveL 198 to (-532.8, -513.42, 952.19) mm, rotated rx 149.35 ry 33.54 rz -64.1 deg; joints [-28.678, -21.072, 36.988, -13.612, 62.219, 0.131, -33.04]
  MoveL 199 to (-494.06, -513.42, 930.04) mm, rotated rx 149.35 ry 33.54 rz -64.1 deg; joints [-28.642, -22.787, 39.005, -14.014, 62.5, 0.473, -33.04]
  MoveL 200 to (-455.86, -513.42, 907) mm, rotated rx 149.35 ry 33.54 rz -64.1 deg; joints [-28.602, -24.499, 41.014, -14.411, 62.782, 0.808, -33.04]
  MoveL 201 to (-418.28, -513.42, 882.95) mm, rotated rx 149.35 ry 33.54 rz -64.1 deg; joints [-28.559, -26.2, 43.015, -14.812, 63.073, 1.142, -33.04]
  MoveL 202 to (-381.55, -513.42, 857.89) mm, rotated rx 149.35 ry 33.54 rz -64.1 deg; joints [-28.512, -27.877, 45.002, -15.228, 63.379, 1.484, -33.04]
  MoveL 203 to (-345.76, -513.42, 831.75) mm, rotated rx 149.35 ry 33.54 rz -64.1 deg; joints [-28.459, -29.523, 46.975, -15.668, 63.708, 1.843, -33.04]
  MoveL 204 to (-314.11, -513.42, 807) mm, rotated rx 149.35 ry 33.54 rz -64.1 deg; joints [-28.405, -30.985, 48.757, -16.099, 64.034, 2.191, -33.04]
  MoveL 205 to (-283.33, -513.42, 781.26) mm, rotated rx 149.35 ry 33.54 rz -64.1 deg; joints [-28.344, -32.406, 50.529, -16.57, 64.394, 2.57, -33.04]
  MoveL 206 to (-253.47, -513.42, 754.49) mm, rotated rx 149.35 ry 33.54 rz -64.1 deg; joints [-28.276, -33.78, 52.291, -17.091, 64.796, 2.986, -33.04]
  MoveL 207 to (-224.56, -513.42, 726.64) mm, rotated rx 163.14 ry 44.09 rz -42.56 deg; joints [-32.78, -37.601, 57.608, -26.32, 48.349, 7.862, -33.04]
  MoveL 208 to (-196.62, -513.42, 697.69) mm, rotated rx 162.55 ry 46.6 rz -44.46 deg; joints [-30.825, -37.995, 60.084, -36.188, 58.754, 10.127, -33.04]
  MoveL 209 to (-169.68, -513.41, 667.6) mm, rotated rx 161.8 ry 49.16 rz -46.66 deg; joints [-28.72, -37.819, 62.447, -45.533, 69.707, 11.196, -33.04]
  MoveL 210 to (-143.76, -513.42, 636.4) mm, rotated rx -172.47 ry 53.81 rz -16.01 deg; joints [-35.203, -40.241, 66.55, -63.162, 60.486, 17.594, -33.04]
  Set speed (1000.0 mm/s)
  MoveL 211 to (-143.76, -513.42, 636.4) mm, rotated rx -172.47 ry 53.81 rz -16.01 deg; joints [-35.203, -40.241, 66.55, -63.162, 60.486, 17.594, -33.04]
  MoveL 212 to (-70.48, -548.09, 694.95) mm, rotated rx -172.47 ry 53.81 rz -16.01 deg; joints [-33.329, -51.45, 67.814, -42.441, 43.539, 7.598, -33.04]
  Set speed (1000.0 mm/s)
  MoveL 213 to (-47.33, -481.42, 695.34) mm, rotated rx 159.13 ry 33.45 rz -61.67 deg; joints [-28.24, -45.438, 58.516, -9.181, 62.09, -12.887, -33.04]
  MoveL 214 to (-103.12, -452.99, 617.38) mm, rotated rx 159.13 ry 33.45 rz -61.67 deg; joints [-30.271, -38.474, 58.619, -15.757, 63.787, -4.136, -33.04]
  MoveL 215 to (-103.12, -452.99, 617.38) mm, rotated rx 159.13 ry 33.45 rz -61.67 deg; joints [-30.271, -38.474, 58.619, -15.757, 63.787, -4.136, -33.04]
  Set speed (50.0 mm/s)
  MoveL 216 to (-129.63, -452.99, 647.84) mm, rotated rx 159.46 ry 32.42 rz -60.95 deg; joints [-31.139, -37.612, 56.614, -11.317, 59.8, -5.914, -33.04]
  MoveL 217 to (-157.02, -452.99, 677.33) mm, rotated rx 159.79 ry 31.39 rz -60.25 deg; joints [-31.935, -36.598, 54.586, -6.876, 56.029, -7.838, -33.04]
  MoveL 218 to (-185.27, -452.99, 705.85) mm, rotated rx 160.11 ry 30.37 rz -59.59 deg; joints [-32.662, -35.458, 52.538, -2.411, 52.449, -9.918, -33.04]
  MoveL 219 to (-214.36, -452.99, 733.45) mm, rotated rx 160.44 ry 29.34 rz -58.94 deg; joints [-33.323, -34.213, 50.473, 2.092, 49.041, -12.161, -33.04]
  MoveL 220 to (-244.27, -452.99, 760.14) mm, rotated rx 160.77 ry 28.31 rz -58.33 deg; joints [-33.921, -32.88, 48.394, 6.648, 45.791, -14.573, -33.04]
  MoveL 221 to (-274.41, -452.99, 785.51) mm, rotated rx 161.11 ry 27.29 rz -57.74 deg; joints [-34.461, -31.499, 46.334, 11.259, 42.685, -17.147, -33.04]
  MoveL 222 to (-305.25, -452.99, 810.1) mm, rotated rx 153.74 ry 18.56 rz -77.17 deg; joints [-30.62, -26.126, 40.435, -0.493, 73.404, -13.225, -33.04]
  MoveL 223 to (-336.79, -452.99, 833.9) mm, rotated rx 154.42 ry 17.71 rz -76.57 deg; joints [-31.073, -24.721, 38.309, 2.176, 71.615, -14.981, -33.04]
  MoveL 224 to (-368.96, -453, 857.01) mm, rotated rx 155.1 ry 16.86 rz -76 deg; joints [-31.48, -23.261, 36.157, 4.742, 70.014, -16.782, -33.04]
  MoveL 225 to (-404.17, -453, 882.18) mm, rotated rx 155.78 ry 16.03 rz -75.46 deg; joints [-31.839, -21.661, 33.813, 7.235, 68.609, -18.708, -33.04]
  MoveL 226 to (-439.94, -453, 906.27) mm, rotated rx 156.47 ry 15.2 rz -74.95 deg; joints [-32.155, -20.015, 31.452, 9.602, 67.397, -20.653, -33.04]
  MoveL 227 to (-476.31, -453, 929.21) mm, rotated rx 157.17 ry 14.38 rz -74.46 deg; joints [-32.431, -18.322, 29.073, 11.835, 66.371, -22.605, -33.04]
  MoveL 228 to (-513.31, -453, 950.92) mm, rotated rx 158.03 ry 13.49 rz -73.96 deg; joints [-32.688, -16.54, 26.603, 14.089, 65.495, -24.788, -33.04]
  MoveL 229 to (-550.97, -453, 971.36) mm, rotated rx 158.59 ry 12.77 rz -73.58 deg; joints [-32.872, -14.798, 24.252, 15.873, 64.864, -26.492, -33.04]
  MoveL 230 to (-589.32, -453, 990.48) mm, rotated rx 159.32 ry 11.98 rz -73.19 deg; joints [-33.041, -12.967, 21.806, 17.667, 64.371, -28.41, -33.04]
  MoveL 231 to (-628.38, -453, 1008.24) mm, rotated rx 160.05 ry 11.21 rz -72.82 deg; joints [-33.18, -11.091, 19.333, 19.305, 64.045, -30.306, -33.04]
  MoveL 232 to (-664.81, -453, 1023.29) mm, rotated rx 160.76 ry 10.39 rz -72.45 deg; joints [-33.338, -9.324, 17.001, 20.987, 63.721, -32.184, -33.04]
  MoveL 233 to (-701.87, -453, 1037.14) mm, rotated rx 162.46 ry 9.16 rz -71.92 deg; joints [-33.495, -7.196, 14.161, 22.931, 63.912, -35.396, -33.04]
  MoveL 234 to (-739.57, -453, 1049.77) mm, rotated rx 164.18 ry 7.94 rz -71.45 deg; joints [-33.615, -5.001, 11.257, 24.556, 64.428, -38.561, -33.04]
  MoveL 235 to (-777.69, -453, 1061.07) mm, rotated rx 165.9 ry 6.74 rz -71.06 deg; joints [-33.698, -2.752, 8.305, 25.839, 65.255, -41.646, -33.04]
  MoveL 236 to (-815.99, -453, 1070.98) mm, rotated rx 167.62 ry 5.56 rz -70.73 deg; joints [-33.747, -0.466, 5.322, 26.781, 66.362, -44.63, -33.04]
  MoveL 237 to (-854.43, -453, 1079.52) mm, rotated rx 169.34 ry 4.43 rz -70.47 deg; joints [-33.766, 1.856, 2.305, 27.399, 67.722, -47.521, -33.04]
  MoveL 238 to (-900.78, -453, 1087.97) mm, rotated rx 171.4 ry 3.13 rz -70.24 deg; joints [-33.754, 4.69, -1.366, 27.739, 69.649, -50.878, -33.04]
  MoveL 239 to (-947.34, -453, 1094.5) mm, rotated rx 173.45 ry 1.9 rz -70.08 deg; joints [-33.707, 7.575, -5.096, 27.674, 71.852, -54.123, -33.04]
  MoveL 240 to (-994.13, -453, 1099.1) mm, rotated rx 175.51 ry 0.75 rz -70 deg; joints [-33.63, 10.515, -8.894, 27.242, 74.29, -57.284, -33.04]
  MoveL 241 to (-1041.13, -453, 1101.84) mm, rotated rx 177.6 ry 0.53 rz -49.99 deg; joints [-36.072, 9.806, -7.417, 67.04, 38.997, -78.938, -33.04]
  MoveL 242 to (-1088.35, -453, 1102.7) mm, rotated rx 179.2 ry -1.1 rz -49.99 deg; joints [-35.854, 12.798, -11.311, 64.962, 42.987, -80.75, -33.04]
  MoveL 243 to (-1134.94, -453, 1101.72) mm, rotated rx -179.2 ry -2.62 rz -50.05 deg; joints [-35.628, 15.797, -15.224, 62.78, 46.942, -82.533, -33.04]
  MoveL 244 to (-1181.72, -453, 1098.96) mm, rotated rx -177.57 ry -4.06 rz -50.15 deg; joints [-35.394, 18.863, -19.243, 60.486, 50.92, -84.351, -33.04]
  MoveL 245 to (-1228.42, -453, 1094.44) mm, rotated rx -175.93 ry -5.41 rz -50.28 deg; joints [-35.153, 21.989, -23.363, 58.106, 54.896, -86.219, -33.04]
  MoveL 246 to (-1274.93, -453, 1088.2) mm, rotated rx -174.27 ry -6.67 rz -50.44 deg; joints [-34.907, 25.18, -27.599, 55.655, 58.86, -88.151, -33.04]
  Set speed (1000.0 mm/s)
  MoveL 247 to (-1274.93, -453, 1088.2) mm, rotated rx -174.27 ry -6.67 rz -50.44 deg; joints [-34.907, 25.18, -27.599, 55.655, 58.86, -88.151, -33.04]
  MoveL 248 to (-1289.99, -450.45, 1187.03) mm, rotated rx -174.27 ry -6.67 rz -50.44 deg; joints [-34.929, 26.223, -32.676, 53.244, 63.693, -91.018, -33.04]
  Set speed (1000.0 mm/s)
  MoveL 249 to (-1255.42, -331.41, 1189.89) mm, rotated rx -175.11 ry -4.63 rz -50.22 deg; joints [-38.135, 24.154, -29.471, 60.413, 55.333, -92.348, -33.04]
  MoveL 250 to (-1243.73, -332.14, 1090.58) mm, rotated rx -175.11 ry -4.63 rz -50.22 deg; joints [-38.165, 23.385, -24.764, 62.958, 50.412, -89.891, -33.04]
  MoveL 251 to (-1243.73, -332.14, 1090.58) mm, rotated rx -175.11 ry -4.63 rz -50.22 deg; joints [-38.165, 23.385, -24.764, 62.958, 50.412, -89.891, -33.04]
  Set speed (50.0 mm/s)
  MoveL 252 to (-1201.21, -332.15, 1094.93) mm, rotated rx -176.65 ry -3.73 rz -50.14 deg; joints [-38.536, 20.631, -21.12, 65.782, 46.768, -88.717, -33.04]
  MoveL 253 to (-1158.6, -332.15, 1097.96) mm, rotated rx -178.19 ry -2.77 rz -50.07 deg; joints [-38.914, 17.921, -17.55, 68.73, 43.002, -87.689, -33.04]
  MoveL 254 to (-1116.04, -332.15, 1099.62) mm, rotated rx -179.13 ry -1.53 rz -70.03 deg; joints [-36.795, 18.924, -19.528, 29.457, 75.984, -66.765, -33.04]
  MoveL 255 to (-1073.65, -332.15, 1099.95) mm, rotated rx 179.1 ry -1.01 rz -69.99 deg; joints [-37.103, 16.233, -16.048, 31.062, 73.295, -64.446, -33.04]
  MoveL 256 to (-1031.4, -332.15, 1098.89) mm, rotated rx 177.31 ry -0.43 rz -69.96 deg; joints [-37.409, 13.588, -12.643, 32.546, 70.635, -62.144, -33.04]
  MoveL 257 to (-989.29, -332.15, 1096.44) mm, rotated rx 175.53 ry 0.22 rz -69.96 deg; joints [-37.715, 10.985, -9.302, 33.9, 68.013, -59.843, -33.04]
  MoveL 258 to (-943.54, -332.15, 1092.18) mm, rotated rx 173.58 ry 0.98 rz -69.98 deg; joints [-38.048, 8.188, -5.721, 35.213, 65.21, -57.321, -33.04]
  MoveL 259 to (-897.97, -332.15, 1086.25) mm, rotated rx 171.63 ry 1.82 rz -70.05 deg; joints [-38.378, 5.43, -2.197, 36.335, 62.485, -54.768, -33.04]
  MoveL 260 to (-852.58, -332.15, 1078.61) mm, rotated rx 169.68 ry 2.72 rz -70.16 deg; joints [-38.706, 2.708, 1.279, 37.244, 59.857, -52.162, -33.04]
  MoveL 261 to (-807.39, -332.15, 1069.24) mm, rotated rx 167.72 ry 3.68 rz -70.32 deg; joints [-39.031, 0.018, 4.712, 37.912, 57.35, -49.481, -33.04]
  MoveL 262 to (-762.39, -332.14, 1058.13) mm, rotated rx 165.76 ry 4.69 rz -70.53 deg; joints [-39.352, -2.639, 8.108, 38.309, 54.997, -46.708, -33.04]
  MoveL 263 to (-717.61, -332.14, 1045.24) mm, rotated rx 163.81 ry 5.74 rz -70.81 deg; joints [-39.667, -5.262, 11.466, 38.403, 52.828, -43.823, -33.04]
  MoveL 264 to (-673.51, -332.14, 1030.7) mm, rotated rx 161.86 ry 6.83 rz -71.15 deg; joints [-39.972, -7.829, 14.761, 38.163, 50.897, -40.831, -33.04]
  MoveL 265 to (-630.2, -332.14, 1014.58) mm, rotated rx 159.94 ry 7.92 rz -71.56 deg; joints [-40.265, -10.331, 17.985, 37.57, 49.235, -37.729, -33.04]
  MoveL 266 to (-587.66, -332.14, 996.91) mm, rotated rx 158.04 ry 9.02 rz -72.03 deg; joints [-40.544, -12.769, 21.141, 36.613, 47.864, -34.509, -33.04]
  MoveL 267 to (-545.88, -332.14, 977.73) mm, rotated rx 156.17 ry 10.11 rz -72.56 deg; joints [-40.81, -15.145, 24.235, 35.29, 46.801, -31.171, -33.04]
  MoveL 268 to (-504.84, -332.14, 957.06) mm, rotated rx 154.31 ry 11.18 rz -73.15 deg; joints [-41.062, -17.458, 27.268, 33.61, 46.053, -27.72, -33.04]
  MoveL 269 to (-464.54, -332.14, 934.92) mm, rotated rx 152.48 ry 12.23 rz -73.79 deg; joints [-41.301, -19.708, 30.244, 31.606, 45.616, -24.178, -33.04]
  MoveL 270 to (-424.95, -332.14, 911.35) mm, rotated rx 150.68 ry 13.23 rz -74.47 deg; joints [-41.532, -21.895, 33.163, 29.337, 45.462, -20.579, -33.04]
  MoveL 271 to (-386.07, -332.14, 886.39) mm, rotated rx 148.92 ry 14.17 rz -75.19 deg; joints [-41.764, -24.02, 36.028, 26.882, 45.546, -16.968, -33.04]
  MoveL 272 to (-348.62, -332.14, 860.6) mm, rotated rx 147.22 ry 15.03 rz -75.9 deg; joints [-42.004, -26.044, 38.783, 24.396, 45.792, -13.47, -33.04]
  MoveL 273 to (-311.87, -332.14, 834.46) mm, rotated rx 148.04 ry 15.08 rz -75.86 deg; joints [-42.273, -27.469, 40.519, 24.341, 45.743, -13.966, -33.04]
  MoveL 274 to (-275.97, -332.14, 805.58) mm, rotated rx 145.2 ry 4 rz -92.77 deg; joints [-40.167, -25.442, 38.126, 14.185, 73.606, -9.252, -33.04]
  MoveL 275 to (-240.89, -332.14, 776.62) mm, rotated rx 145.2 ry 4 rz -92.77 deg; joints [-40.592, -26.947, 40.163, 14.634, 72.698, -8.793, -33.04]
  MoveL 276 to (-197.3, -332.14, 738.58) mm, rotated rx 145.2 ry 4 rz -92.77 deg; joints [-41.166, -28.819, 42.735, 15.227, 71.486, -8.198, -33.04]
  MoveL 277 to (-154.73, -332.14, 699.38) mm, rotated rx 145.2 ry 4 rz -92.77 deg; joints [-41.782, -30.652, 45.284, 15.85, 70.206, -7.601, -33.04]
  MoveL 278 to (-112.95, -332.14, 659.29) mm, rotated rx 145.2 ry 4 rz -92.77 deg; joints [-42.45, -32.461, 47.814, 16.515, 68.849, -7.018, -33.04]
  MoveL 279 to (-71.68, -332.14, 618.61) mm, rotated rx 145.2 ry 4 rz -92.77 deg; joints [-43.182, -34.27, 50.329, 17.243, 67.402, -6.479, -33.04]
  MoveL 280 to (-45.8, -332.14, 590.77) mm, rotated rx 145.2 ry 4 rz -92.77 deg; joints [-43.68, -35.376, 51.961, 17.713, 66.409, -6.065, -33.04]
  Set speed (1000.0 mm/s)
  MoveL 281 to (-45.8, -332.14, 590.77) mm, rotated rx 145.2 ry 4 rz -92.77 deg; joints [-43.68, -35.376, 51.961, 17.713, 66.409, -6.065, -33.04]
  MoveL 282 to (10.93, -340.62, 672.69) mm, rotated rx 145.2 ry 4 rz -92.77 deg; joints [-44.432, -41.037, 51.577, 20.159, 67.35, -12.957, -33.04]
  Set speed (1000.0 mm/s)
  MoveL 283 to (38.13, -274.14, 652.27) mm, rotated rx 136.01 ry 1 rz -90.96 deg; joints [-57.418, -44.842, 55.932, 53.324, 34.043, -17.049, -33.04]
  MoveL 284 to (-31.3, -271.71, 580.34) mm, rotated rx 136.01 ry 1 rz -90.96 deg; joints [-54.279, -38.304, 55.568, 42.395, 38.217, -5.487, -33.04]
  MoveL 285 to (-31.3, -271.71, 580.34) mm, rotated rx 136.01 ry 1 rz -90.96 deg; joints [-54.279, -38.304, 55.568, 42.395, 38.217, -5.487, -33.04]
  Set speed (50.0 mm/s)
  MoveL 286 to (-72.29, -271.71, 623.84) mm, rotated rx 137.02 ry 1.5 rz -91.39 deg; joints [-51.942, -36.204, 52.644, 36.486, 44.556, -4.457, -33.04]
  MoveL 287 to (-114, -271.71, 666.47) mm, rotated rx 137.34 ry 1.99 rz -91.84 deg; joints [-50.007, -34.263, 49.986, 31.909, 49.491, -3.466, -33.04]
  MoveL 288 to (-156.65, -271.71, 707.95) mm, rotated rx 138.06 ry 2.49 rz -92.23 deg; joints [-48.231, -32.157, 47.162, 27.992, 54.102, -3.381, -33.04]
  MoveL 289 to (-200.42, -271.71, 748.07) mm, rotated rx 138.34 ry 2.79 rz -92.48 deg; joints [-46.889, -30.155, 44.483, 25.434, 57.315, -3.425, -33.04]
  MoveL 290 to (-235.68, -271.71, 778.54) mm, rotated rx 139.9 ry 2.69 rz -92.27 deg; joints [-46.129, -28.242, 41.836, 24.937, 59.24, -5.629, -33.04]
  MoveL 291 to (-271.77, -271.71, 808) mm, rotated rx 141.56 ry 2.52 rz -92 deg; joints [-45.47, -26.269, 39.119, 24.681, 60.986, -8.036, -33.04]
  MoveL 292 to (-308.73, -271.71, 836.39) mm, rotated rx 143.31 ry 2.28 rz -91.7 deg; joints [-44.882, -24.229, 36.335, 24.541, 62.661, -10.58, -33.04]
  MoveL 293 to (-346.61, -271.71, 863.66) mm, rotated rx 145.13 ry 2 rz -91.39 deg; joints [-44.342, -22.121, 33.481, 24.429, 64.339, -13.221, -33.04]
  MoveL 294 to (-386.26, -271.71, 890.29) mm, rotated rx 147.07 ry 1.67 rz -91.08 deg; joints [-43.826, -19.897, 30.497, 24.279, 66.11, -15.986, -33.04]
  MoveL 295 to (-426.95, -271.72, 915.64) mm, rotated rx 149.07 ry 1.31 rz -90.78 deg; joints [-43.333, -17.596, 27.438, 24.041, 67.979, -18.801, -33.04]
  MoveL 296 to (-468.73, -271.72, 939.66) mm, rotated rx 151.12 ry 0.93 rz -90.52 deg; joints [-42.857, -15.217, 24.3, 23.68, 69.972, -21.657, -33.04]
  MoveL 297 to (-511.36, -271.72, 962.16) mm, rotated rx 153.23 ry 0.55 rz -90.28 deg; joints [-42.395, -12.773, 21.1, 23.168, 72.096, -24.528, -33.04]
  MoveL 298 to (-554.58, -271.71, 982.98) mm, rotated rx 155.35 ry 0.18 rz -90.08 deg; joints [-41.946, -10.28, 17.857, 22.49, 74.345, -27.391, -33.04]
  MoveL 299 to (-598.41, -271.72, 1002.09) mm, rotated rx 158.67 ry 7.35 rz -71.35 deg; joints [-43.877, -11.427, 19.6, 46.91, 40.752, -40.445, -33.04]
  MoveL 300 to (-642.81, -271.72, 1019.52) mm, rotated rx 160.62 ry 6.34 rz -70.98 deg; joints [-43.352, -8.897, 16.33, 46.614, 43.15, -43.154, -33.04]
  MoveL 301 to (-687.81, -271.72, 1035.24) mm, rotated rx 162.58 ry 5.34 rz -70.68 deg; joints [-42.836, -6.318, 13.009, 46.036, 45.727, -45.755, -33.04]
  MoveL 302 to (-733.4, -271.72, 1049.25) mm, rotated rx 164.55 ry 4.38 rz -70.43 deg; joints [-42.329, -3.689, 9.635, 45.205, 48.455, -48.269, -33.04]
  MoveL 303 to (-779.59, -271.72, 1061.55) mm, rotated rx 166.54 ry 3.45 rz -70.24 deg; joints [-41.83, -1.009, 6.202, 44.148, 51.31, -50.719, -33.04]
  MoveL 304 to (-826.38, -271.72, 1072.13) mm, rotated rx 168.54 ry 2.57 rz -70.1 deg; joints [-41.339, 1.724, 2.706, 42.889, 54.271, -53.125, -33.04]
  MoveL 305 to (-873.78, -271.72, 1080.96) mm, rotated rx 170.55 ry 1.74 rz -70.01 deg; joints [-40.854, 4.513, -0.86, 41.445, 57.317, -55.503, -33.04]
  MoveL 306 to (-921.52, -271.72, 1088.01) mm, rotated rx 172.56 ry 0.97 rz -69.96 deg; joints [-40.379, 7.343, -4.481, 39.843, 60.412, -57.859, -33.04]
  MoveL 307 to (-969.31, -271.72, 1093.25) mm, rotated rx 174.56 ry 0.28 rz -69.94 deg; joints [-39.914, 10.203, -8.146, 38.111, 63.523, -60.197, -33.04]
  MoveL 308 to (-1013.17, -271.72, 1096.5) mm, rotated rx 176.39 ry -0.29 rz -69.95 deg; joints [-39.496, 12.855, -11.551, 36.42, 66.379, -62.34, -33.04]
  MoveL 309 to (-1057.07, -271.72, 1098.31) mm, rotated rx 178.21 ry -0.79 rz -69.97 deg; joints [-39.087, 15.54, -15.009, 34.643, 69.228, -64.491, -33.04]
  MoveL 310 to (-1101.01, -271.72, 1098.68) mm, rotated rx -179.99 ry -1.22 rz -70 deg; joints [-38.684, 18.263, -18.53, 32.785, 72.065, -66.665, -33.04]
  MoveL 311 to (-1144.98, -271.72, 1097.65) mm, rotated rx -178.19 ry -1.58 rz -70.04 deg; joints [-38.288, 21.031, -22.128, 30.854, 74.885, -68.875, -33.04]
  MoveL 312 to (-1189, -271.72, 1095.25) mm, rotated rx -177.26 ry -2.99 rz -50.09 deg; joints [-40.316, 20.116, -20.201, 70.571, 42.336, -90.462, -33.04]
  MoveL 313 to (-1233.06, -271.72, 1091.47) mm, rotated rx -175.66 ry -3.8 rz -50.15 deg; joints [-39.862, 22.892, -23.888, 67.214, 46.212, -91.291, -33.04]
  Set speed (1000.0 mm/s)
  MoveL 314 to (-1233.06, -271.72, 1091.47) mm, rotated rx -175.66 ry -3.8 rz -50.15 deg; joints [-39.862, 22.892, -23.888, 67.214, 46.212, -91.291, -33.04]
  MoveL 315 to (-1243.1, -271.49, 1190.96) mm, rotated rx -175.66 ry -3.8 rz -50.15 deg; joints [-39.819, 23.548, -28.453, 64.478, 51.262, -93.5, -33.04]
  Set speed (1000.0 mm/s)
  MoveL 316 to (-1233.53, -211.37, 1191.81) mm, rotated rx -176.28 ry -3.06 rz -50.1 deg; joints [-41.534, 23.184, -27.751, 68.913, 47.201, -94.987, -33.04]
  MoveL 317 to (-1225.12, -211.3, 1092.15) mm, rotated rx -175.46 ry -1.61 rz -70.06 deg; joints [-39.182, 26.378, -29.025, 29.68, 76.883, -73.163, -33.04]
  MoveL 318 to (-1225.12, -211.3, 1092.15) mm, rotated rx -175.46 ry -1.61 rz -70.06 deg; joints [-39.182, 26.378, -29.025, 29.68, 76.883, -73.163, -33.04]
  Set speed (50.0 mm/s)
  MoveL 319 to (-1180.77, -211.29, 1095.25) mm, rotated rx -177.2 ry -1.49 rz -70.05 deg; joints [-39.634, 23.546, -25.288, 31.871, 74.107, -71.045, -33.04]
  MoveL 320 to (-1136.43, -211.29, 1097.03) mm, rotated rx -178.95 ry -1.29 rz -70.02 deg; joints [-40.097, 20.772, -21.653, 34.032, 71.279, -68.99, -33.04]
  MoveL 321 to (-1092.13, -211.29, 1097.45) mm, rotated rx 179.28 ry -1.03 rz -69.99 deg; joints [-40.57, 18.049, -18.102, 36.161, 68.4, -66.992, -33.04]
  MoveL 322 to (-1047.86, -211.29, 1096.51) mm, rotated rx 177.5 ry -0.7 rz -69.96 deg; joints [-41.055, 15.367, -14.622, 38.257, 65.472, -65.04, -33.04]
  MoveL 323 to (-1003.63, -211.29, 1094.18) mm, rotated rx 175.71 ry -0.29 rz -69.93 deg; joints [-41.554, 12.722, -11.2, 40.319, 62.496, -63.128, -33.04]
  MoveL 324 to (-959.44, -211.29, 1090.44) mm, rotated rx 173.91 ry 0.18 rz -69.91 deg; joints [-42.067, 10.106, -7.826, 42.348, 59.473, -61.246, -33.04]
  MoveL 325 to (-911.27, -211.29, 1084.68) mm, rotated rx 171.93 ry 0.77 rz -69.91 deg; joints [-42.646, 7.283, -4.189, 44.52, 56.123, -59.222, -33.04]
  MoveL 326 to (-863.35, -211.29, 1077.19) mm, rotated rx 169.95 ry 1.43 rz -69.94 deg; joints [-43.243, 4.499, -0.605, 46.64, 52.738, -57.228, -33.04]
  MoveL 327 to (-815.97, -211.29, 1067.99) mm, rotated rx 167.97 ry 2.15 rz -70 deg; joints [-43.858, 1.766, 2.913, 48.695, 49.342, -55.267, -33.04]
  MoveL 328 to (-769.14, -211.29, 1057.1) mm, rotated rx 166 ry 2.93 rz -70.11 deg; joints [-44.491, -0.916, 6.373, 50.685, 45.939, -53.333, -33.04]
  MoveL 329 to (-722.85, -211.29, 1044.51) mm, rotated rx 164.04 ry 3.75 rz -70.25 deg; joints [-45.147, -3.552, 9.781, 52.612, 42.533, -51.42, -33.04]
  MoveL 330 to (-677.11, -211.29, 1030.23) mm, rotated rx 162.08 ry 4.62 rz -70.44 deg; joints [-45.827, -6.14, 13.14, 54.481, 39.129, -49.524, -33.04]
  MoveL 331 to (-631.9, -211.29, 1014.26) mm, rotated rx 159.46 ry -1.46 rz -89.45 deg; joints [-44.046, -5.042, 11.269, 26.255, 73.723, -34.48, -33.04]
  MoveL 332 to (-587.26, -211.29, 996.59) mm, rotated rx 157.34 ry -1.2 rz -89.5 deg; joints [-44.662, -7.61, 14.589, 27.791, 70.795, -31.907, -33.04]
  MoveL 333 to (-543.15, -211.29, 977.22) mm, rotated rx 155.23 ry -0.92 rz -89.58 deg; joints [-45.302, -10.134, 17.868, 29.207, 67.921, -29.344, -33.04]
  MoveL 334 to (-499.58, -211.29, 956.14) mm, rotated rx 153.13 ry -0.62 rz -89.69 deg; joints [-45.971, -12.613, 21.109, 30.508, 65.103, -26.788, -33.04]
  MoveL 335 to (-456.71, -211.29, 933.44) mm, rotated rx 151.05 ry -0.31 rz -89.83 deg; joints [-46.67, -15.039, 24.302, 31.7, 62.346, -24.248, -33.04]
  MoveL 336 to (-414.9, -211.29, 909.34) mm, rotated rx 149.02 ry 0 rz -90 deg; joints [-47.398, -17.389, 27.421, 32.789, 59.666, -21.748, -33.04]
  MoveL 337 to (-374.18, -211.29, 883.92) mm, rotated rx 147.04 ry 0.31 rz -90.2 deg; joints [-48.158, -19.662, 30.468, 33.798, 57.05, -19.295, -33.04]
  MoveL 338 to (-334.49, -211.29, 857.23) mm, rotated rx 145.12 ry 0.6 rz -90.42 deg; joints [-48.958, -21.86, 33.447, 34.755, 54.476, -16.896, -33.04]
  MoveL 339 to (-296.56, -211.29, 829.88) mm, rotated rx 143.28 ry 0.86 rz -90.64 deg; joints [-49.789, -23.939, 36.302, 35.68, 51.967, -14.612, -33.04]
  MoveL 340 to (-259.56, -211.29, 801.39) mm, rotated rx 141.51 ry 1.09 rz -90.87 deg; joints [-50.678, -25.945, 39.096, 36.645, 49.429, -12.416, -33.04]
  MoveL 341 to (-223.46, -211.29, 771.8) mm, rotated rx 139.8 ry 1.28 rz -91.08 deg; joints [-51.64, -27.878, 41.831, 37.72, 46.807, -10.345, -33.04]
  MoveL 342 to (-188.21, -211.29, 741.16) mm, rotated rx 138.16 ry 1.42 rz -91.27 deg; joints [-52.695, -29.735, 44.508, 39.01, 44.018, -8.454, -33.04]
  MoveL 343 to (-153.17, -211.29, 708.92) mm, rotated rx 136.58 ry 1.5 rz -91.42 deg; joints [-53.897, -31.546, 47.174, 40.711, 40.881, -6.81, -33.04]
  MoveL 344 to (-118.94, -211.29, 675.68) mm, rotated rx 135.08 ry 1.51 rz -91.5 deg; joints [-55.271, -33.274, 49.783, 43.081, 37.24, -5.616, -33.04]
  MoveL 345 to (-85.47, -211.29, 641.51) mm, rotated rx 133.7 ry 1.41 rz -91.47 deg; joints [-56.884, -34.914, 52.337, 46.615, 32.752, -5.176, -33.04]
  MoveL 346 to (-52.71, -211.28, 606.47) mm, rotated rx 132.45 ry 1.18 rz -91.29 deg; joints [-58.833, -36.456, 54.851, 52.356, 26.737, -6.151, -33.04]
  MoveL 347 to (-20.57, -211.28, 570.66) mm, rotated rx 131.36 ry 0.78 rz -90.89 deg; joints [-61.276, -37.885, 57.395, 63.468, 17.243, -10.531, -33.04]
  Set speed (1000.0 mm/s)
  MoveL 348 to (-20.57, -211.28, 570.66) mm, rotated rx 131.36 ry 0.78 rz -90.89 deg; joints [-61.276, -37.885, 57.395, 63.468, 17.243, -10.531, -33.04]
  MoveL 349 to (54.46, -213.35, 636.73) mm, rotated rx 132.94 ry -14.11 rz -104.36 deg; joints [-62.699, -41.082, 53.291, 56.837, 45.777, -12.219, -33.04]
  Set speed (1000.0 mm/s)
  MoveL 350 to (64.02, -151.87, 627.18) mm, rotated rx 132.16 ry -14.71 rz -103.72 deg; joints [-68.488, -39.237, 53.387, 73.355, 31.687, -20.161, -33.04]
  MoveL 351 to (-12.03, -150.86, 562.25) mm, rotated rx 132.16 ry -14.71 rz -103.72 deg; joints [-64.682, -33.322, 52.736, 65.277, 33.554, -9.751, -33.04]
  MoveL 352 to (-12.03, -150.86, 562.25) mm, rotated rx 132.16 ry -14.71 rz -103.72 deg; joints [-64.682, -33.322, 52.736, 65.277, 33.554, -9.751, -33.04]
  Set speed (50.0 mm/s)
  MoveL 353 to (-43.87, -150.86, 598.66) mm, rotated rx 133.5 ry -14.28 rz -104.17 deg; joints [-62.683, -32, 50.176, 58.572, 40.152, -8.121, -33.04]
  MoveL 354 to (-76.48, -150.86, 634.15) mm, rotated rx 133.3 ry 0.52 rz -90.55 deg; joints [-63.02, -33.398, 52.566, 77.041, 9.38, -21.219, -33.04]
  MoveL 355 to (-109.89, -150.86, 668.68) mm, rotated rx 134.82 ry 0.47 rz -90.47 deg; joints [-61.192, -31.939, 49.755, 65.693, 18.883, -17.023, -33.04]
  MoveL 356 to (-144.14, -150.86, 702.21) mm, rotated rx 136.42 ry 0.37 rz -90.35 deg; joints [-59.567, -30.357, 47.034, 59.808, 24.934, -16.169, -33.04]
  MoveL 357 to (-179.28, -150.86, 734.69) mm, rotated rx 138.07 ry 0.23 rz -90.2 deg; joints [-58.093, -28.664, 44.3, 55.738, 29.804, -16.46, -33.04]
  MoveL 358 to (-214.66, -150.86, 765.54) mm, rotated rx 139.76 ry 0.05 rz -90.04 deg; joints [-56.76, -26.901, 41.578, 52.629, 33.99, -17.332, -33.04]
  MoveL 359 to (-250.95, -150.86, 795.32) mm, rotated rx 141.5 ry -0.15 rz -89.88 deg; joints [-55.522, -25.048, 38.811, 50.03, 37.824, -18.561, -33.04]
  MoveL 360 to (-288.17, -150.86, 823.99) mm, rotated rx 143.29 ry -0.38 rz -89.72 deg; joints [-54.362, -23.107, 35.993, 47.744, 41.436, -20.034, -33.04]
  MoveL 361 to (-326.35, -150.86, 851.52) mm, rotated rx 145.13 ry -0.62 rz -89.56 deg; joints [-53.271, -21.084, 33.12, 45.652, 44.908, -21.684, -33.04]
  MoveL 362 to (-366.33, -150.86, 878.38) mm, rotated rx 147.06 ry -0.88 rz -89.43 deg; joints [-52.218, -18.936, 30.127, 43.635, 48.364, -23.509, -33.04]
  MoveL 363 to (-407.38, -150.86, 903.99) mm, rotated rx 149.03 ry -1.15 rz -89.31 deg; joints [-51.218, -16.706, 27.069, 41.678, 51.771, -25.449, -33.04]
  MoveL 364 to (-449.53, -150.86, 928.26) mm, rotated rx 151.06 ry -1.42 rz -89.22 deg; joints [-50.265, -14.394, 23.941, 39.739, 55.16, -27.487, -33.04]
  MoveL 365 to (-492.48, -150.86, 951.01) mm, rotated rx 153.11 ry -1.67 rz -89.15 deg; joints [-49.361, -12.018, 20.764, 37.799, 58.526, -29.596, -33.04]
  MoveL 366 to (-536.02, -150.86, 972.1) mm, rotated rx 155.17 ry -1.91 rz -89.11 deg; joints [-48.504, -9.594, 17.551, 35.842, 61.869, -31.754, -33.04]
  MoveL 367 to (-580.13, -150.86, 991.54) mm, rotated rx 157.25 ry -2.13 rz -89.11 deg; joints [-47.69, -7.121, 14.299, 33.848, 65.201, -33.96, -33.04]
  MoveL 368 to (-624.83, -150.86, 1009.32) mm, rotated rx 159.33 ry -2.32 rz -89.13 deg; joints [-46.913, -4.6, 11.006, 31.804, 68.526, -36.208, -33.04]
  MoveL 369 to (-670.11, -150.86, 1025.45) mm, rotated rx 161.41 ry -2.47 rz -89.17 deg; joints [-46.17, -2.034, 7.667, 29.696, 71.85, -38.497, -33.04]
  MoveL 370 to (-715.96, -150.86, 1039.94) mm, rotated rx 163.49 ry -2.58 rz -89.24 deg; joints [-45.457, 0.581, 4.28, 27.512, 75.178, -40.83, -33.04]
  MoveL 371 to (-762.42, -150.86, 1052.79) mm, rotated rx 165.52 ry 2.41 rz -69.96 deg; joints [-47.074, -0.515, 6.257, 57.708, 40.528, -56.545, -33.04]
  MoveL 372 to (-809.44, -150.86, 1063.98) mm, rotated rx 167.47 ry 1.72 rz -69.9 deg; joints [-46.312, 2.119, 2.811, 54.853, 44.438, -57.911, -33.04]
  MoveL 373 to (-857.05, -150.86, 1073.53) mm, rotated rx 169.42 ry 1.08 rz -69.86 deg; joints [-45.577, 4.805, -0.69, 52.094, 48.236, -59.395, -33.04]
  MoveL 374 to (-905.11, -150.86, 1081.4) mm, rotated rx 171.37 ry 0.52 rz -69.86 deg; joints [-44.871, 7.537, -4.244, 49.401, 51.93, -60.977, -33.04]
  MoveL 375 to (-953.28, -150.86, 1087.55) mm, rotated rx 173.3 ry 0.02 rz -69.88 deg; joints [-44.193, 10.299, -7.835, 46.767, 55.507, -62.637, -33.04]
  MoveL 376 to (-997.51, -150.86, 1091.74) mm, rotated rx 175.06 ry -0.36 rz -69.9 deg; joints [-43.595, 12.859, -11.165, 44.388, 58.69, -64.221, -33.04]
  MoveL 377 to (-1041.8, -150.86, 1094.55) mm, rotated rx 176.81 ry -0.67 rz -69.94 deg; joints [-43.017, 15.449, -14.541, 42.032, 61.787, -65.865, -33.04]
  MoveL 378 to (-1086.16, -150.86, 1096.03) mm, rotated rx 178.55 ry -0.91 rz -69.98 deg; joints [-42.457, 18.075, -17.971, 39.689, 64.803, -67.569, -33.04]
  MoveL 379 to (-1130.58, -150.86, 1096.2) mm, rotated rx -179.73 ry -1.09 rz -70.01 deg; joints [-41.914, 20.742, -21.469, 37.355, 67.74, -69.336, -33.04]
  MoveL 380 to (-1175.06, -150.86, 1095.07) mm, rotated rx -178.02 ry -1.18 rz -70.03 deg; joints [-41.385, 23.458, -25.048, 35.025, 70.6, -71.172, -33.04]
  MoveL 381 to (-1219.6, -150.87, 1092.68) mm, rotated rx -176.32 ry -1.21 rz -70.03 deg; joints [-40.87, 26.231, -28.724, 32.695, 73.384, -73.081, -33.04]
  Set speed (1000.0 mm/s)
  MoveL 382 to (-1219.6, -150.87, 1092.68) mm, rotated rx -176.32 ry -1.21 rz -70.03 deg; joints [-40.87, 26.231, -28.724, 32.695, 73.384, -73.081, -33.04]
  MoveL 383 to (-1226.34, -151.09, 1192.44) mm, rotated rx -176.32 ry -1.21 rz -70.03 deg; joints [-40.828, 26.808, -33.172, 31.218, 77.016, -76.671, -33.04]
  Set speed (1000.0 mm/s)
  MoveL 384 to (-1219.95, -90.54, 1192.95) mm, rotated rx -177.94 ry -0.68 rz -70.01 deg; joints [-42.611, 26.371, -32.437, 35.075, 72.679, -75.906, -33.04]
  MoveL 385 to (-1216.16, -90.44, 1093.02) mm, rotated rx -177.94 ry -0.68 rz -70.01 deg; joints [-42.633, 25.959, -28.213, 36.422, 69.102, -72.437, -33.04]
  MoveL 386 to (-1216.16, -90.44, 1093.02) mm, rotated rx -177.94 ry -0.68 rz -70.01 deg; joints [-42.633, 25.959, -28.213, 36.422, 69.102, -72.437, -33.04]
  Set speed (50.0 mm/s)
  MoveL 387 to (-1162.45, -90.44, 1094.89) mm, rotated rx -179.55 ry -0.06 rz -70 deg; joints [-43.114, 22.681, -23.735, 38.378, 65.819, -70.116, -33.04]
  MoveL 388 to (-1108.8, -90.44, 1095.01) mm, rotated rx 178.76 ry 0.61 rz -70.01 deg; joints [-43.627, 19.484, -19.413, 40.328, 62.51, -67.839, -33.04]
  MoveL 389 to (-1055.22, -90.44, 1093.33) mm, rotated rx 177.01 ry 1.29 rz -70.04 deg; joints [-44.178, 16.363, -15.232, 42.294, 59.179, -65.632, -33.04]
  MoveL 390 to (-1001.7, -90.44, 1089.8) mm, rotated rx 175.21 ry 2 rz -70.09 deg; joints [-44.77, 13.304, -11.163, 44.299, 55.802, -63.488, -33.04]
  MoveL 391 to (-948.26, -90.44, 1084.35) mm, rotated rx 173.35 ry 2.72 rz -70.18 deg; joints [-45.409, 10.295, -7.184, 46.369, 52.352, -61.407, -33.04]
  MoveL 392 to (-899.86, -90.44, 1077.71) mm, rotated rx 171.61 ry 3.38 rz -70.27 deg; joints [-46.033, 7.604, -3.636, 48.329, 49.138, -59.577, -33.04]
  MoveL 393 to (-851.97, -90.44, 1069.49) mm, rotated rx 169.84 ry 4.06 rz -70.4 deg; joints [-46.698, 4.968, -0.166, 50.377, 45.85, -57.829, -33.04]
  MoveL 394 to (-804.61, -90.44, 1059.68) mm, rotated rx 168.04 ry 4.74 rz -70.54 deg; joints [-47.406, 2.384, 3.236, 52.546, 42.465, -56.177, -33.04]
  MoveL 395 to (-757.78, -90.44, 1048.27) mm, rotated rx 166.21 ry 5.42 rz -70.71 deg; joints [-48.163, -0.151, 6.58, 54.882, 38.951, -54.644, -33.04]
  MoveL 396 to (-711.48, -90.44, 1035.25) mm, rotated rx 163.24 ry 0.47 rz -90.14 deg; joints [-46.487, 0.99, 4.591, 24.817, 74.026, -38.916, -33.04]
  MoveL 397 to (-665.74, -90.44, 1020.64) mm, rotated rx 161.26 ry 0.5 rz -90.17 deg; joints [-47.233, -1.529, 7.883, 26.829, 70.934, -36.612, -33.04]
  MoveL 398 to (-620.52, -90.44, 1004.41) mm, rotated rx 159.27 ry 0.53 rz -90.2 deg; joints [-48.03, -4.005, 11.126, 28.875, 67.776, -34.372, -33.04]
  MoveL 399 to (-575.85, -90.44, 986.56) mm, rotated rx 157.27 ry 0.56 rz -90.24 deg; joints [-48.883, -6.436, 14.327, 30.972, 64.536, -32.201, -33.04]
  MoveL 400 to (-531.73, -90.44, 967.08) mm, rotated rx 155.26 ry 0.59 rz -90.27 deg; joints [-49.798, -8.823, 17.49, 33.14, 61.2, -30.108, -33.04]
  MoveL 401 to (-488.15, -90.43, 945.96) mm, rotated rx 153.25 ry 0.62 rz -90.31 deg; joints [-50.779, -11.163, 20.618, 35.401, 57.753, -28.108, -33.04]
  MoveL 402 to (-445.12, -90.43, 923.19) mm, rotated rx 151.24 ry 0.64 rz -90.35 deg; joints [-51.834, -13.455, 23.715, 37.787, 54.169, -26.219, -33.04]
  MoveL 403 to (-402.74, -90.43, 898.81) mm, rotated rx 149.25 ry 0.66 rz -90.39 deg; joints [-52.967, -15.69, 26.779, 40.337, 50.425, -24.466, -33.04]
  MoveL 404 to (-361.43, -90.43, 873.08) mm, rotated rx 147.29 ry 0.67 rz -90.43 deg; joints [-54.174, -17.843, 29.781, 43.079, 46.523, -22.9, -33.04]
  MoveL 405 to (-321.19, -90.43, 846.09) mm, rotated rx 145.37 ry 0.68 rz -90.47 deg; joints [-55.458, -19.909, 32.725, 46.083, 42.418, -21.562, -33.04]
  MoveL 406 to (-282.77, -90.43, 818.44) mm, rotated rx 143.54 ry 0.69 rz -90.51 deg; joints [-56.798, -21.845, 35.558, 49.387, 38.13, -20.535, -33.04]
  MoveL 407 to (-245.34, -90.43, 789.64) mm, rotated rx 141.75 ry 0.69 rz -90.54 deg; joints [-58.228, -23.69, 38.347, 53.216, 33.471, -19.887, -33.04]
  MoveL 408 to (-208.84, -90.43, 759.73) mm, rotated rx 140 ry 0.68 rz -90.57 deg; joints [-59.756, -25.437, 41.102, 57.866, 28.259, -19.798, -33.04]
  MoveL 409 to (-173.27, -90.43, 728.73) mm, rotated rx 138.3 ry 0.66 rz -90.59 deg; joints [-61.395, -27.08, 43.842, 63.971, 22.102, -20.65, -33.04]
  MoveL 410 to (-137.98, -90.43, 696.08) mm, rotated rx 136.61 ry 0.64 rz -90.6 deg; joints [-63.195, -28.633, 46.678, 73.735, 13.598, -23.724, -33.04]
  MoveL 411 to (-103.59, -90.43, 662.36) mm, rotated rx 136.6 ry -13.42 rz -104.99 deg; joints [-62.826, -27.269, 44.332, 55.166, 44.284, -10.671, -33.04]
  MoveL 412 to (-70.09, -90.43, 627.6) mm, rotated rx 135.03 ry -13.85 rz -104.59 deg; joints [-64.665, -28.709, 46.981, 60.908, 38.245, -11.354, -33.04]
  MoveL 413 to (-37.45, -90.43, 591.83) mm, rotated rx 133.51 ry -14.28 rz -104.17 deg; joints [-66.628, -30.005, 49.612, 68.058, 31.316, -13.032, -33.04]
  MoveL 414 to (-5.64, -90.43, 555.08) mm, rotated rx 132.04 ry -14.71 rz -103.71 deg; joints [-68.714, -31.134, 52.259, 77.939, 22.722, -16.531, -33.04]
  Set speed (1000.0 mm/s)
  MoveL 415 to (-5.64, -90.43, 555.08) mm, rotated rx 132.04 ry -14.71 rz -103.71 deg; joints [-68.714, -31.134, 52.259, 77.939, 22.722, -16.531, -33.04]
  MoveL 416 to (70.54, -91.52, 619.84) mm, rotated rx 132.04 ry -14.71 rz -103.71 deg; joints [-72.592, -36.801, 53.024, 89.473, 19.1, -29.043, -33.04]
  Set speed (1000.0 mm/s)
  MoveL 417 to (74.94, -30.36, 613.76) mm, rotated rx 137.81 ry -29.25 rz -118.6 deg; joints [-75.821, -30.361, 46.882, 74.411, 45.973, -20.609, -33.04]
  MoveL 418 to (-1.36, -30, 549.12) mm, rotated rx 137.81 ry -29.25 rz -118.6 deg; joints [-72.229, -25.547, 46.454, 72.356, 44.429, -13.837, -33.04]
  MoveL 419 to (-1.36, -30, 549.12) mm, rotated rx 137.81 ry -29.25 rz -118.6 deg; joints [-72.229, -25.547, 46.454, 72.356, 44.429, -13.837, -33.04]
  Set speed (50.0 mm/s)
  MoveL 420 to (-33.27, -30, 585.93) mm, rotated rx 133.51 ry -14.63 rz -103.79 deg; joints [-70.504, -27.717, 48.947, 83.765, 19.144, -22.052, -33.04]
  MoveL 421 to (-66.03, -30, 621.75) mm, rotated rx 135.05 ry -14.24 rz -104.19 deg; joints [-68.533, -26.614, 46.246, 72.683, 28.38, -17.849, -33.04]
  MoveL 422 to (-99.65, -30, 656.55) mm, rotated rx 136.63 ry -13.84 rz -104.58 deg; joints [-66.63, -25.347, 43.58, 64.892, 35.636, -15.796, -33.04]
  MoveL 423 to (-134.15, -30.01, 690.3) mm, rotated rx 138.26 ry -13.42 rz -104.97 deg; joints [-64.815, -23.934, 40.9, 58.676, 41.927, -14.843, -33.04]
  MoveL 424 to (-169.57, -30.01, 722.98) mm, rotated rx 139.93 ry -12.98 rz -105.35 deg; joints [-63.092, -22.391, 38.189, 53.394, 47.623, -14.593, -33.04]
  MoveL 425 to (-205.26, -30.01, 754.01) mm, rotated rx 139.92 ry 0.21 rz -90.17 deg; joints [-63.576, -23.77, 40.685, 76.169, 14.534, -29.796, -33.04]
  MoveL 426 to (-241.87, -30.01, 783.95) mm, rotated rx 141.67 ry 0.21 rz -90.17 deg; joints [-61.905, -22.154, 37.821, 66.552, 22.815, -26.81, -33.04]
  MoveL 427 to (-279.43, -30.01, 812.78) mm, rotated rx 143.46 ry 0.21 rz -90.16 deg; joints [-60.33, -20.427, 34.993, 60.172, 29.087, -25.86, -33.04]
  MoveL 428 to (-317.96, -30.01, 840.46) mm, rotated rx 145.29 ry 0.21 rz -90.14 deg; joints [-58.845, -18.597, 32.146, 55.22, 34.452, -25.851, -33.04]
  MoveL 429 to (-358.31, -30.01, 867.49) mm, rotated rx 147.2 ry 0.21 rz -90.13 deg; joints [-57.418, -16.628, 29.199, 51.011, 39.376, -26.43, -33.04]
  MoveL 430 to (-399.74, -30.01, 893.25) mm, rotated rx 149.15 ry 0.2 rz -90.12 deg; joints [-56.072, -14.563, 26.2, 47.35, 43.925, -27.42, -33.04]
  MoveL 431 to (-442.21, -30.01, 917.67) mm, rotated rx 151.14 ry 0.2 rz -90.11 deg; joints [-54.805, -12.406, 23.143, 44.069, 48.203, -28.716, -33.04]
  MoveL 432 to (-485.33, -30.01, 940.5) mm, rotated rx 153.14 ry 0.19 rz -90.1 deg; joints [-53.623, -10.186, 20.055, 41.09, 52.233, -30.235, -33.04]
  MoveL 433 to (-529.01, -30.01, 961.7) mm, rotated rx 155.14 ry 0.19 rz -90.09 deg; joints [-52.52, -7.909, 16.936, 38.338, 56.062, -31.927, -33.04]
  MoveL 434 to (-573.23, -30.01, 981.28) mm, rotated rx 157.14 ry 0.18 rz -90.07 deg; joints [-51.492, -5.578, 13.781, 35.756, 59.729, -33.76, -33.04]
  MoveL 435 to (-618, -30.01, 999.25) mm, rotated rx 159.13 ry 0.17 rz -90.06 deg; joints [-50.531, -3.198, 10.588, 33.305, 63.257, -35.708, -33.04]
  MoveL 436 to (-663.3, -30.01, 1015.63) mm, rotated rx 161.11 ry 0.16 rz -90.05 deg; joints [-49.633, -0.77, 7.353, 30.956, 66.667, -37.753, -33.04]
  MoveL 437 to (-709.14, -30.01, 1030.42) mm, rotated rx 163.07 ry 0.15 rz -90.05 deg; joints [-48.792, 1.707, 4.067, 28.682, 69.98, -39.884, -33.04]
  MoveL 438 to (-755.51, -30.01, 1043.64) mm, rotated rx 165.02 ry 0.14 rz -90.04 deg; joints [-48.004, 4.233, 0.724, 26.462, 73.214, -42.095, -33.04]
  MoveL 439 to (-802.41, -30.01, 1055.31) mm, rotated rx 167.75 ry 4.56 rz -70.5 deg; joints [-49.635, 3.107, 2.788, 58.457, 37.717, -58.963, -33.04]
  MoveL 440 to (-849.83, -30.01, 1065.43) mm, rotated rx 169.53 ry 3.91 rz -70.37 deg; joints [-48.842, 5.648, -0.619, 55.631, 41.519, -60.2, -33.04]
  MoveL 441 to (-897.78, -30.01, 1074.01) mm, rotated rx 171.28 ry 3.27 rz -70.26 deg; joints [-48.098, 8.243, -4.092, 53.056, 45.142, -61.611, -33.04]
  MoveL 442 to (-946.21, -30.01, 1081.06) mm, rotated rx 173 ry 2.64 rz -70.17 deg; joints [-47.4, 10.894, -7.64, 50.666, 48.631, -63.16, -33.04]
  MoveL 443 to (-999.71, -30.01, 1087.03) mm, rotated rx 174.84 ry 1.96 rz -70.09 deg; joints [-46.684, 13.861, -11.621, 48.208, 52.328, -64.982, -33.04]
  MoveL 444 to (-1053.3, -30.01, 1091.16) mm, rotated rx 176.62 ry 1.31 rz -70.04 deg; joints [-46.021, 16.883, -15.692, 45.885, 55.909, -66.906, -33.04]
  MoveL 445 to (-1106.98, -30.01, 1093.53) mm, rotated rx 178.33 ry 0.67 rz -70.01 deg; joints [-45.403, 19.969, -19.879, 43.655, 59.407, -68.924, -33.04]
  MoveL 446 to (-1160.73, -30.01, 1094.19) mm, rotated rx 179.99 ry 0.05 rz -70 deg; joints [-44.828, 23.134, -24.21, 41.484, 62.856, -71.034, -33.04]
  MoveL 447 to (-1214.57, -30.01, 1093.19) mm, rotated rx -178.41 ry -0.55 rz -70.01 deg; joints [-44.289, 26.397, -28.722, 39.341, 66.284, -73.239, -33.04]
  Set speed (1000.0 mm/s)
  MoveL 448 to (-1214.57, -30.01, 1093.19) mm, rotated rx -178.41 ry -0.55 rz -70.01 deg; joints [-44.289, 26.397, -28.722, 39.341, 66.284, -73.239, -33.04]
  MoveL 449 to (-1217.5, -30.06, 1193.15) mm, rotated rx -178.41 ry -0.55 rz -70.01 deg; joints [-44.273, 26.78, -32.912, 38.001, 69.915, -76.636, -33.04]

